(* Logix 5000 project; controller CIP_14485201 vendor 1 type 14 code 216 rev 38.11; software revision 38.01 *)

TASK MainProgram (periodic, rate 20 ms, priority 1, watchdog 40 ms) : MainProgram
TASK PID_SupplyFlow (periodic, rate 250 ms, priority 5, watchdog 500 ms) : PID_SupplyFlow

MODULES
   Local : vendor 1 type 14 code 216 (5069 0, rev 38.11)
        Module:7:I.1   // SPARE IN-426
        Module:7:I.6   // SPARE IN-436
        Module:7:I.7   // SPARE IN-438
        Module:7:I.0   // CHEM #1 TANK LOW LEVEL LSL-201
        Module:7:I.2   // CHEM #2 TANK LOW LEVEL LSL-301
        Module:7:I.3   // SPARE IN-430
        Module:7:I.4   // SPARE IN-432
        Module:7:I.5   // SPARE IN-434
        Module:7:I   // 8-PT DIG. INPUT
        Module:9:O.7   // SPARE OUT-396
        Module:9:O.0   // AIR BLOW BLOCK XY-008
        Module:9:O.2   // CHEM #1 ENABLE XY-202
        Module:9:O.3   // CHEM #2 ENABLE XY-302
        Module:9:O.5   // CHEM #2 BLOCK XY-305
        Module:9:O.6   // OVERFLOW TANK DRAIN PUMP XV-032
        Module:9:O.4   // CHEM #1 BLOCK XY-205
        Module:9:O.1   // SPARE OUT-384
        Module:9:O   // 8-PT DIG. OUTPUT
        Module:10:I   // 8-PT DIG. OUTPUT
        Module:10:O.1   // LOW POINT DRAIN XY-023
        Module:10:O.3   // SPARE SOLENOID SV-410
        Module:10:O.4   // SPARE SOLENOID SV-412
        Module:10:O.0   // OVERFLOW TANK DRAIN XY-022
        Module:10:O.2   // DRAIN TO WASTE NEUTRALIZATION XY-024
        Module:10:O.5   // SPARE OUT-414
        Module:10:O.6   // SPARE OUT-416
        Module:10:O.7   // SPARE OUT-418
        Module:10:O   // 8-PT DIG. OUTPUT
        Module:6:I.7   // SPARE IN-356
        Module:6:I.0   // SEP. TANK HIGH LEVEL LSH-101
        Module:6:I.1   // SUPPLY PUMP FAULT CONTACT JY-001C
        Module:6:I.2   // SEP. TANK MIDDLE LEVEL LSM-110
        Module:6:I.3   // HEATER CONTACTOR ALARM CONTACT JY-004B
        Module:6:I.4   // HEATER HIGH TEMP CONTACT TSH-004
        Module:6:I.5   // DRAIN PUMP LOW LEVEL LSL-405
        Module:6:I.6   // OVERFLOW TANK HIGH LEVEL LSH-401
        Module:6:I   // 8-PT DIG. INPUT
        Module:5:I.5   // SPARE IN-334
        Module:5:I.6   // SPARE IN-336
        Module:5:I.0   // CONTROL POWER ON CP-153
        Module:5:I.1   // LOCAL E-STOP PRESSED PBLT-125
        Module:5:I.2   // SEPARATOR TANK BURST SENSOR PSH-106
        Module:5:I.3   // AIR SUPPLY PRESSURE PSL-021
        Module:5:I.4   // SUPPLY PUMP AUX CONTACT JY-001B
        Module:5:I.7   // SEP. TANK LOW LEVEL LSL-105
        Module:5:I   // 8-PT DIG. INPUT
        Module:8:O.1   // AIR BLOW XV-008A
        Module:8:O.6   // ALARM HORN AH-376
        Module:8:O.5   // RETURN TO DRAIN XY-018
        Module:8:O.4   // SPARE SOLENOID SV-372
        Module:8:O.7   // HEATER ENABLE JY-004A
        Module:8:O.0   // SEP. TANK AWFI FILL XY-102
        Module:8:O.2   // SUPPLY PUMP CASING DRAIN XY-002
        Module:8:O.3   // SUPPLY PUMP ENABLE JY-001A
        Module:8:O   // 8-PT DIG. OUTPUT
        Module:8:I   // 8-PT DIG. OUTPUT
        Module:9:I.4   // SPARE IN-432
        Module:9:I.5   // SPARE IN-434
        Module:9:I.6   // SPARE IN-436
        Module:9:I.7   // SPARE IN-438
        Module:9:I.0   // CHEM 1 TANK LOW LEVEL LSL-201
        Module:9:I.1   // CHEM 1 TANK HIGH LEVEL LSH-201
        Module:9:I.2   // CHEM 2 TANK LOW LEVEL LSL-301
        Module:9:I.3   // CHEM 2 TANK HIGH LEVEL LSH-301
        Module:9:I   // 8-PT DIG. OUTPUT
      Module : 1734-AENT (Ethernet 192.168.1.50, rev 4.1, Output RPI 20 ms)
         Analog_In1 : vendor 1 type 115 code 210 (PointIO 1, rev 3.1, Input RPI 80 ms)
              Module:1:C   // 8-PT ANALOG INPUT
              Module:1:I.Ch2Data   // RINSE CONDUCTIVITY 0-10 uS/cm AE-019
              Module:1:I.Ch3Data   // WASH CONDUCTIVITY 0-100 mS/cm AE-104
              Module:1:I.Ch0Data   // SUPPLY TEMPERATURE 0-100°C TT-005
              Module:1:I.Ch1Data   // RETURN TEMPERATURE 0-100°C TT-017
              Module:1:I.Ch2Fault   // RINSE CONDUCTIVITY 0-10 uS/cm AE-019 FAULT
              Module:1:I.Ch2Underrange   // RINSE CONDUCTIVITY 0-10 uS/cm AE-019 UNDERRANGE
              Module:1:I.Ch1Underrange   // RETURN TEMPERATURE 0-100°C TT-017 UNDERRANGE
              Module:1:I.Ch1Overrange   // RETURN TEMPERATURE 0-100°C TT-017 OVERRANGE
              Module:1:I.Ch0Overrange   // SUPPLY TEMPERATURE 0-100°C TT-005 OVERRANGE
              Module:1:I.Ch1Fault   // RETURN TEMPERATURE 0-100°C TT-017 FAULT
              Module:1:I.Ch6Data   // SUPPLY PRESSURE 0-100 PSIG PIT-009
              Module:1:I.Ch7Data   // SPARE IN-272
              Module:1:I.Ch4Data   // SUPPLY FLOW 0-60 GPM FIT-010
              Module:1:I.Ch5Data   // SPARE IN-264
              Module:1:I.Ch0Fault   // SUPPLY TEMPERATURE 0-100°C TT-005 FAULT
              Module:1:I.Ch0Underrange   // SUPPLY TEMPERATURE 0-100°C TT-005 UNDERRANGE
              Module:1:I.Ch2Overrange   // RINSE CONDUCTIVITY 0-10 uS/cm AE-019 OVERRANGE
              Module:1:I.Ch3Fault   // WASH CONDUCTIVITY 0-100 mS/cm AE-104 FAULT
              Module:1:I.Ch3Underrange   // WASH CONDUCTIVITY 0-100 mS/cm AE-104 UNDERRANGE
              Module:1:I.Ch3Overrange   // WASH CONDUCTIVITY 0-100 mS/cm AE-104 OVERRANGE
              Module:1:I.Ch4Fault   // SUPPLY FLOW 0-60 GPM FIT-010 FAULT
              Module:1:I.Ch4Underrange   // SUPPLY FLOW 0-60 GPM FIT-010 UNDERRANGE
              Module:1:I.Ch4Overrange   // SUPPLY FLOW 0-60 GPM FIT-010 OVERRANGE
              Module:1:I.Ch5Fault   // SPARE IN-264 FAULT
              Module:1:I.Ch5Underrange   // SPARE IN-264 UNDERRANGE
              Module:1:I.Ch5Overrange   // SPARE IN-264 OVERRANGE
              Module:1:I.Ch6Fault   // SUPPLY PRESSURE 0-100 PSIG PIT-009 FAULT
              Module:1:I.Ch6Underrange   // SUPPLY PRESSURE 0-100 PSIG PIT-009 UNDERRANGE
              Module:1:I.Ch6Overrange   // SUPPLY PRESSURE 0-100 PSIG PIT-009 OVERRANGE
              Module:1:I.Ch7Fault   // SPARE IN-272 FAULT
              Module:1:I.Ch7Underrange   // SPARE IN-272 UNDERRANGE
              Module:1:I.Ch7Overrange   // SPARE IN-272 OVERRANGE
              Module:1:I   // 8-PT ANALOG INPUT
         Analog_In2 : 1734-IE2C (PointIO 2, rev 3.1, Input RPI 80 ms)
              Module:2:C   // 2-PT ANALOG OUTPUT
              Module:2:I.Ch1Fault   // DRAIN FLOW FEEDBACK POSTION 0-100% FY-006B FAULT
              Module:2:I.Ch1Overrange   // DRAIN FLOW FEEDBACK POSTION 0-100% FY-006B OVERRANGE
              Module:2:I.Ch0Fault   // SUPPLY FLOW FEEDBACK POSTION 0-100% FY-003B FAULT
              Module:2:I.Ch0Overrange   // SUPPLY FLOW FEEDBACK POSTION 0-100% FY-003B OVERRANGE
              Module:2:I.Ch0Underrange   // SUPPLY FLOW FEEDBACK POSTION 0-100% FY-003B UNDERRANGE
              Module:2:I.Ch1Underrange   // DRAIN FLOW FEEDBACK POSTION 0-100% FY-006B UNDERRANGE
              Module:2:I.Ch0Data   // SUPPLY FLOW FEEDBACK POSTION 0-100% FY-003B
              Module:2:I.Ch1Data   // DRAIN FLOW FEEDBACK POSTION 0-100% FY-006B
              Module:2:I   // 2-PT ANALOG OUTPUT
         Discrete_In3 : 1734-IB8 (PointIO 7, rev 3.1)
              Module:7:C   // 8-PT DIG. INPUT
         Discrete_In1 : 1734-IB8 (PointIO 5, rev 3.1)
              Module:5:C   // 8-PT DIG. INPUT
         Discrete_In2 : 1734-IB8 (PointIO 6, rev 3.1)
              Module:6:C   // 8-PT DIG. INPUT
         Discrete_Out2 : 1734-OB8 (PointIO 9, rev 3.1)
              Module:9:C   // 8-PT DIG. OUTPUT
         Analog_Out1 : 1734-OE2C (PointIO 3, rev 3.1, Output RPI 80 ms)
              Module:3:C   // 2-PT ANALOG OUTPUT
              Module:3:I.Ch0Fault   // SUPPLY FLOW FEEDBACK POSTION 0-100% FY-003B FAULT
              Module:3:I.Ch1Fault   // DRAIN FLOW FEEDBACK POSTION 0-100% FY-006B FAULT
              Module:3:I   // 2-PT ANALOG OUTPUT
              Module:3:O.Ch0Data   // SPARE OUT-284
              Module:3:O.Ch1Data   // SUPPLY FLOW MODULATION 0-100% FY-003A
              Module:3:O   // 2-PT ANALOG OUTPUT
         Analog_Out2 : 1734-OE2C (PointIO 4, rev 3.1, Output RPI 80 ms)
              Module:4:C   // 8-PT DIG. INPUT
              Module:4:I   // 8-PT DIG. INPUT
              Module:4:O.Ch0Data   // DRAIN FLOW MODULATION 0-100% FY-006A
              Module:4:O.Ch1Data   // SPARE OUT-298
              Module:4:O   // 2-PT ANALOG OUTPUT
         Discrete_Out1 : 1734-OB8 (PointIO 8, rev 3.1)
              Module:8:C   // 8-PT DIG. OUTPUT
         Discrete_Out3 : 1734-OB8 (PointIO 10, rev 3.1)
              Module:10:C   // 8-PT DIG. OUTPUT
END_MODULES

TYPE CIP_to_Process :
STRUCT
   DINT : DINT[4];
   REAL : REAL[20];
   STRING : STRING[5];
END_STRUCT
END_TYPE

TYPE Process_to_CIP :
STRUCT
   DINT : DINT[2];
   REAL : REAL[2];
END_STRUCT
END_TYPE

TYPE RECIPE :
STRUCT
   OpCode : DINT[97];   // OPCODES
   StepTime : DINT[97];   // STEP TIMES
   Setpoint : REAL[97];   // SETPOINTS
   Name : STRING;   // NAME
END_STRUCT
END_TYPE

TYPE Wash_Control :
STRUCT
   Print_Control : DINT;   // PRINT CONTROL
   Print_Control_One_Shot : DINT;   // ONE SHOT
   Print_Control_String : STRING[3];   // PRINT CONTROL STRING
   Timer : TIMER[4];   // PRINT RATE TO ASCII PORT
END_STRUCT
END_TYPE

TYPE Wash_Data :
STRUCT
   Start_Time : STRING;   // START TIME
   Stop_Time : STRING;   // STOP TIME
   Required_Time : DINT[6];   // REQUIRED TIME
   Required_Time_String : STRING[6];   // REQUIRED TIME STRING
   Temperature : DINT[3];   // TEMPERATURE
   Temperature_String : STRING[6];   // TEMPERATURE STRING
   Conductivity : DINT[3];   // CONDUCTIVITY
   Conductivity_String : STRING[6];   // CONDUCTIVITY STRING
   Flow : DINT[3];   // SUPPLY FLOW
   Flow_String : STRING[6];   // SUPPLY FLOW STRING
   Pressure : DINT[3];   // SUPPLY PRESSURE
   Pressure_String : STRING[6];   // SUPPLY PRESSURE STRING
   Sample_Timer : TIMER;   // SAMPLE TIMER
   Counter : COUNTER;   // SAMPLE COUNTER
   Print_Text : STRING[3];   // PRINT SPACE
   Active : BOOL[32];   // ACTIVE
END_STRUCT
END_TYPE

TYPE Wash_Data_Control :
STRUCT
   Control : DINT[2];   // DATA CONTROL
   One_Shot : DINT;   // DATA CONTROL ONE SHOT
   Print_Active_Pin : BOOL;   // PRINT ACTIVE PIN FROM OPCODE PINNING CHART
   Timer : TIMER;   // PRINT WASH DELAY CLEAR ALLOW FOR DATA TO BE TRANSFERED TO THE TABLE
END_STRUCT
END_TYPE

TYPE Wash_Steps :
STRUCT
   Wash_Steps : STRING[40];
   Print_Step : DINT[2];
END_STRUCT
END_TYPE

VAR_GLOBAL   (* controller tags *)
   Alarm_Ack : INT[8];   // ALARMS ACKNOWLEDGE BITS
        [2].15   // ALARM 47 ACKNOWLEDGE
        [2].2   // ALARM 34 ACKNOWLEDGE
        [2].13   // ALARM 45 ACKNOWLEDGE
        [2].14   // ALARM 46 ACKNOWLEDGE
        [6].0   // ALARM 96 ACKNOWLEDGE
        [6].1   // ALARM 97 ACKNOWLEDGE
        [6].2   // ALARM 98 ACKNOWLEDGE
        [6].10   // ALARM 106 ACKNOWLEDGE
        [6].11   // ALARM 107 ACKNOWLEDGE
        [6].12   // ALARM 108 ACKNOWLEDGE
        [6].13   // ALARM 109 ACKNOWLEDGE
        [2].3   // ALARM 35 ACKNOWLEDGE
        [2].4   // ALARM 36 ACKNOWLEDGE
        [2].5   // ALARM 37 ACKNOWLEDGE
        [6].14   // ALARM 110 ACKNOWLEDGE
        [6].15   // ALARM 111 ACKNOWLEDGE
        [2].6   // ALARM 38 ACKNOWLEDGE
        [2].7   // ALARM 39 ACKNOWLEDGE
        [2].8   // ALARM 40 ACKNOWLEDGE
        [6].3   // ALARM 99 ACKNOWLEDGE
        [6].4   // ALARM 100 ACKNOWLEDGE
        [6].5   // ALARM 101 ACKNOWLEDGE
        [2].9   // ALARM 41 ACKNOWLEDGE
        [3]   // ALARMS 48-63 ACKNOWLEDGE BITS
        [6].6   // ALARM 102 ACKNOWLEDGE
        [6].7   // ALARM 103 ACKNOWLEDGE
        [6].8   // ALARM 104 ACKNOWLEDGE
        [3].0   // ALARM 48 ACKNOWLEDGE
        [3].1   // ALARM 49 ACKNOWLEDGE
        [3].2   // ALARM 50 ACKNOWLEDGE
        [6].9   // ALARM 105 ACKNOWLEDGE
        [7]   // ALARMS 97-127 ACKNOWLEDGE BITS
        [3].10   // ALARM 58 ACKNOWLEDGE
        [3].11   // ALARM 59 ACKNOWLEDGE
        [0]   // ALARMS 1-15 ACKNOWLEDGE BITS
        [7].0   // ALARM 112 ACKNOWLEDGE
        [7].1   // ALARM 113 ACKNOWLEDGE
        [7].10   // ALARM 122 ACKNOWLEDGE
        [3].12   // ALARM 60 ACKNOWLEDGE
        [3].13   // ALARM 61 ACKNOWLEDGE
        [0].1   // ALARM 1 ACKNOWLEDGE
        [0].10   // ALARM 10 ACKNOWLEDGE
        [7].11   // ALARM 123 ACKNOWLEDGE
        [7].12   // ALARM 124 ACKNOWLEDGE
        [3].14   // ALARM 62 ACKNOWLEDGE
        [3].15   // ALARM 63 ACKNOWLEDGE
        [0].11   // ALARM 11 ACKNOWLEDGE
        [0].12   // ALARM 12 ACKNOWLEDGE
        [7].13   // ALARM 125 ACKNOWLEDGE
        [7].14   // ALARM 126 ACKNOWLEDGE
        [3].3   // ALARM 51 ACKNOWLEDGE
        [3].4   // ALARM 52 ACKNOWLEDGE
        [3].5   // ALARM 53 ACKNOWLEDGE
        [0].13   // ALARM 13 ACKNOWLEDGE
        [0].14   // ALARM 14 ACKNOWLEDGE
        [7].15   // ALARM 127 ACKNOWLEDGE
        [7].2   // ALARM 114 ACKNOWLEDGE
        [7].3   // ALARM 115 ACKNOWLEDGE
        [3].6   // ALARM 54 ACKNOWLEDGE
        [3].7   // ALARM 55 ACKNOWLEDGE
        [3].8   // ALARM 56 ACKNOWLEDGE
        [0].15   // ALARM 15 ACKNOWLEDGE
        [0].2   // ALARM 2 ACKNOWLEDGE
        [7].4   // ALARM 116 ACKNOWLEDGE
        [7].5   // ALARM 117 ACKNOWLEDGE
        [7].6   // ALARM 118 ACKNOWLEDGE
        [3].9   // ALARM 57 ACKNOWLEDGE
        [4]   // ALARMS 64-79 ACKNOWLEDGE BITS
        [0].3   // ALARM 3 ACKNOWLEDGE
        [0].4   // ALARM 4 ACKNOWLEDGE
        [0].5   // ALARM 5 ACKNOWLEDGE
        [7].7   // ALARM 119 ACKNOWLEDGE
        [7].8   // ALARM 120 ACKNOWLEDGE
        [7].9   // ALARM 121 ACKNOWLEDGE
        [4].0   // ALARM 64 ACKNOWLEDGE
        [4].1   // ALARM 65 ACKNOWLEDGE
        [4].2   // ALARM 66 ACKNOWLEDGE
        [0].6   // ALARM 6 ACKNOWLEDGE
        [0].7   // ALARM 7 ACKNOWLEDGE
        [0].8   // ALARM 8 ACKNOWLEDGE
        [4].10   // ALARM 74 ACKNOWLEDGE
        [4].11   // ALARM 75 ACKNOWLEDGE
        [0].9   // ALARM 9 ACKNOWLEDGE
        [1]   // ALARMS 16-31 ACKNOWLEDGE BITS
        [4].12   // ALARM 76 ACKNOWLEDGE
        [4].13   // ALARM 77 ACKNOWLEDGE
        [1].0   // ALARM 16 ACKNOWLEDGE
        [1].1   // ALARM 17 ACKNOWLEDGE
        [4].14   // ALARM 78 ACKNOWLEDGE
        [4].15   // ALARM 79 ACKNOWLEDGE
        [1].10   // ALARM 26 ACKNOWLEDGE
        [1].11   // ALARM 27 ACKNOWLEDGE
        [4].3   // ALARM 67 ACKNOWLEDGE
        [4].4   // ALARM 68 ACKNOWLEDGE
        [4].5   // ALARM 69 ACKNOWLEDGE
        [1].12   // ALARM 28 ACKNOWLEDGE
        [1].13   // ALARM 29 ACKNOWLEDGE
        [4].6   // ALARM 70 ACKNOWLEDGE
        [4].7   // ALARM 71 ACKNOWLEDGE
        [4].8   // ALARM 72 ACKNOWLEDGE
        [1].14   // ALARM 30 ACKNOWLEDGE
        [1].15   // ALARM 31 ACKNOWLEDGE
        [4].9   // ALARM 73 ACKNOWLEDGE
        [5]   // ALARMS 80-95 ACKNOWLEDGE BITS
        [1].2   // ALARM 18 ACKNOWLEDGE
        [1].3   // ALARM 19 ACKNOWLEDGE
        [5].0   // ALARM 80 ACKNOWLEDGE
        [5].1   // ALARM 81 ACKNOWLEDGE
        [5].2   // ALARM 82 ACKNOWLEDGE
        [1].4   // ALARM 20 ACKNOWLEDGE
        [1].5   // ALARM 21 ACKNOWLEDGE
        [5].10   // ALARM 90 ACKNOWLEDGE
        [5].11   // ALARM 91 ACKNOWLEDGE
        [1].6   // ALARM 22 ACKNOWLEDGE
        [1].7   // ALARM 23 ACKNOWLEDGE
        [5].12   // ALARM 92 ACKNOWLEDGE
        [5].13   // ALARM 93 ACKNOWLEDGE
        [1].8   // ALARM 24 ACKNOWLEDGE
        [1].9   // ALARM 25 ACKNOWLEDGE
        [5].14   // ALARM 94 ACKNOWLEDGE
        [5].15   // ALARM 95 ACKNOWLEDGE
        [2]   // ALARMS 32-47 ACKNOWLEDGE BITS
        [2].0   // ALARM 32 ACKNOWLEDGE
        [5].3   // ALARM 83 ACKNOWLEDGE
        [5].4   // ALARM 84 ACKNOWLEDGE
        [5].5   // ALARM 85 ACKNOWLEDGE
        [2].1   // ALARM 33 ACKNOWLEDGE
        [2].10   // ALARM 42 ACKNOWLEDGE
        [5].6   // ALARM 86 ACKNOWLEDGE
        [5].7   // ALARM 87 ACKNOWLEDGE
        [5].8   // ALARM 88 ACKNOWLEDGE
        [2].11   // ALARM 43 ACKNOWLEDGE
        [2].12   // ALARM 44 ACKNOWLEDGE
        [5].9   // ALARM 89 ACKNOWLEDGE
        [6]   // ALARMS 96-111 ACKNOWLEDGE BITS
   Alarm_Ack_All_PB : BOOL;   // SYSTEM ALARM ACK ALL PUSHBUTTON ON ALARM PAGE
   Alarm_Present : INT[8] := ([0] := 70, [2] := 98);   // ALARM MSGS 1-127 PRESENT BITS
        [7].0   // ALARM 112 PRESENT
        [7].1   // ALARM 113 PRESENT
        [7].10   // ALARM 122 PRESENT
        [1].3   // ALARM 19 SUPPLY TEMPERATURE HOLD WATCHDOG PRESENT
        [1].4   // ALARM 20 RETURN TEMPERATURE HOLD WATCHDOG PRESENT
        [1].15   // ALARM 31 SEPARATOR TANK LOW LEVEL PRESENT
        [1].2   // ALARM 18 SEPARATOR TANK EMPTY HOLD WATCHDOG PRESENT
        [7].11   // ALARM 123 PRESENT
        [7].12   // ALARM 124 PRESENT
        [7].13   // ALARM 125 PRESENT
        [3].0   // ALARM 48 PRESENT
        [3].1   // ALARM 49 PRESENT
        [3].10   // ALARM 58 PRESENT
        [7].14   // ALARM 126 PRESENT
        [7].15   // ALARM 127 PRESENT
        [7].2   // ALARM 114 PRESENT
        [3].11   // ALARM 59 PRESENT
        [3].12   // ALARM 60 PRESENT
        [3].13   // ALARM 61 PRESENT
        [7].3   // ALARM 115 PRESENT
        [7].4   // ALARM 116 PRESENT
        [7].5   // ALARM 117 PRESENT
        [3].14   // ALARM 62 PRESENT
        [3].15   // ALARM 63 PRESENT
        [3].2   // ALARM 50 PRESENT
        [7].6   // ALARM 118 PRESENT
        [7].7   // ALARM 119 PRESENT
        [7].8   // ALARM 120 PRESENT
        [3].3   // ALARM 51 PRESENT
        [3].4   // ALARM 52 PRESENT
        [3].5   // ALARM 53 PRESENT
        [7].9   // ALARM 121 PRESENT
        [3].6   // ALARM 54 PRESENT
        [3].7   // ALARM 55 PRESENT
        [3].8   // ALARM 56 PRESENT
        [3].9   // ALARM 57 PRESENT
        [4]   // ALARM MSGS 64-79 PRESENT BITS
        [4].0   // ALARM 64 PRESENT
        [4].1   // ALARM 65 PRESENT
        [4].10   // ALARM 74 PRESENT
        [4].11   // ALARM 75 PRESENT
        [4].12   // ALARM 76 PRESENT
        [4].13   // ALARM 77 PRESENT
        [4].14   // ALARM 78 PRESENT
        [4].15   // ALARM 79 PRESENT
        [4].2   // ALARM 66 PRESENT
        [4].3   // ALARM 67 PRESENT
        [4].4   // ALARM 68 PRESENT
        [4].5   // ALARM 69 PRESENT
        [4].6   // ALARM 70 PRESENT
        [4].7   // ALARM 71 PRESENT
        [4].8   // ALARM 72 PRESENT
        [4].9   // ALARM 73 PRESENT
        [5]   // ALARM MSGS 80-95 PRESENT BITS
        [5].0   // ALARM 80 PRESENT
        [5].1   // ALARM 81 PRESENT
        [5].10   // ALARM 90 PRESENT
        [5].11   // ALARM 91 PRESENT
        [5].12   // ALARM 92 PRESENT
        [5].13   // ALARM 93 PRESENT
        [0]   // ALARM MSGS 1-15 PRESENT BITS
        [0].0   // ALARM 0 N/A PRESENT
        [5].14   // ALARM 94 PRESENT
        [5].15   // ALARM 95 PRESENT
        [5].2   // ALARM 82 PRESENT
        [0].1   // ALARM 1 LOSS OF CONTROL POWER PRESENT
        [0].10   // ALARM 10 WASH CONDUCTIVITY SENSOR FAILURE PRESENT
        [0].5   // ALARM 5 PRESENT
        [5].3   // ALARM 83 PRESENT
        [5].4   // ALARM 84 PRESENT
        [5].5   // ALARM 85 PRESENT
        [0].11   // ALARM 11 SUPPLY FLOW SENSOR FAILURE PRESENT
        [0].12   // ALARM 12 SUPPLY FLOW FEEDBACK SENSOR FAILURE PRESENT
        [5].6   // ALARM 86 PRESENT
        [5].7   // ALARM 87 PRESENT
        [5].8   // ALARM 88 PRESENT
        [0].13   // ALARM 13 SUPPLY PRESSURE SENSOR FAILURE PRESENT
        [0].14   // ALARM 14 DRAIN FLOW FEEDBACK SENSOR FAILURE PRESENT
        [5].9   // ALARM 89 PRESENT
        [6]   // ALARM MSGS 96-111 PRESENT BITS
        [0].15   // ALARM 15 SUPPLY PUMP FAILURE PRESENT
        [0].2   // ALARM 2 LOSS OF PLC POWER PRESENT
        [6].0   // ALARM 96 PRESENT
        [6].1   // ALARM 97 PRESENT
        [6].10   // ALARM 106 PRESENT
        [0].3   // ALARM 3 LOCAL E-STOP PRESSED PRESENT
        [0].6   // ALARM 6 I/O COMMUNICATION FAILURE PRESENT
        [0].4   // ALARM 4 PRESENT
        [1].5   // ALARM 21 RINSE CONDUCTIVITY HOLD WATCHDOG PRESENT
        [1].6   // ALARM 22 CHEM #1 CONDUCTIVITY HOLD WATCHDOG PRESENT
        [6].11   // ALARM 107 PRESENT
        [6].12   // ALARM 108 PRESENT
        [6].2   // ALARM 98 PRESENT
        [0].7   // ALARM 7 SUPPLY TEMPERATURE SENSOR FAILURE PRESENT
        [0].8   // ALARM 8 RETURN TEMPERATURE SENSOR FAILURE PRESENT
        [1].7   // ALARM 23 CHEM #2 CONDUCTIVITY HOLD WATCHDOG PRESENT
        [1].8   // ALARM 24 OVERFLOW TANK EMPTY HOLD WATCHDOG PRESENT
        [6].13   // ALARM 109 PRESENT
        [6].14   // ALARM 110 PRESENT
        [6].3   // ALARM 99 PRESENT
        [0].9   // ALARM 9 RINSE CONDUCTIVITY SENSOR FAILURE PRESENT
        [1]   // ALARM MSGS 16-31 PRESENT BITS
        [6].15   // ALARM 111 PRESENT
        [6].4   // ALARM 100 PRESENT
        [6].5   // ALARM 101 PRESENT
        [1].1   // ALARM 17 SEPARATOR TANK FILL HOLD WATCHDOG PRESENT
        [1].10   // ALARM 26 HIGH SUPPLY FLOW PRESENT
        [6].6   // ALARM 102 PRESENT
        [6].7   // ALARM 103 PRESENT
        [6].8   // ALARM 104 PRESENT
        [1].11   // ALARM 27 LOW SUPPLY FLOW PRESENT
        [1].12   // ALARM 28 HIGH SUPPLY PRESSURE PRESENT
        [1].0   // ALARM 16 PRESENT
        [6].9   // ALARM 105 PRESENT
        [7]   // ALARM MSGS 112-127 PRESENT BITS
        [1].13   // ALARM 29 LOW SUPPLY PRESSURE PRESENT
        [1].14   // ALARM 30 PRESENT
        [2].0   // ALARM 32 PRESENT
        [1].9   // ALARM 25 HIGH SUPPLY TEMPERATURE PRESENT
        [2]   // ALARM MSGS 32-47 PRESENT BITS
        [2].1   // ALARM 33 HEATER CONTACTOR FAULT PRESENT
        [2].10   // ALARM 42 PRESENT
        [2].11   // ALARM 43 PRESENT
        [2].12   // ALARM 44 PRESENT
        [2].13   // ALARM 45 PRESENT
        [2].14   // ALARM 46 PROCESS EQUIPMENT HEARTBEAT FAILURE PRESENT
        [2].15   // ALARM 47 PROCESS EQUIPMENT STOP ACTIVE PRESENT
        [2].2   // ALARM 34 HEATER ELEMENT HIGH TEMPERATURE PRESENT
        [2].3   // ALARM 35 CHEM #1 TANK LOW LEVEL PRESENT
        [2].4   // ALARM 36 CHEM #2 TANK LOW LEVEL PRESENT
        [2].5   // ALARM 37 PANEL AIR PRESSURE FAILURE PRESENT
        [2].6   // ALARM 38 SEP. TANK BURST SENSOR FAILURE PRESENT
        [2].8   // ALARM 40 SUPPLY FLOW MODULATION VALVE FAILURE PRESENT
        [2].9   // ALARM 41 DRAIN FLOW MODULATION VALVE FAILURE PRESENT
        [3]   // ALARM MSGS 48-63 PRESENT BITS
        [2].7   // ALARM 39 PRESENT
   Alarm_Preset_Indx : DINT := 84;   // ALARM TIMER PRESET INDEX POSITION
   Alarm_Remote_Ack_All : BOOL;   // SYSTEM ALARM ACK ALL TAG USED ON ALARM SETUP ADVANCED TAB TOGGLES EVEYTIME THE ACK_ALL BUTTON IS PUSHED
   Alarm_Status_Reset : BOOL;   // SYSTEM ALARM ACK ALL TAG USED ON ALARM SETUP ADVANCED TAB TOGGLES EVERYTIME THE HISTORY CLEAR ALL IS PUSHED
   Alarm_Timer : TIMER[128] := ([1].ACC := 20, [1].EN := 1, [1].DN := 1, [2].ACC := 20, [2].EN := 1, [2].DN := 1, [6].PRE := 3000, [7].PRE := 5000, [8].PRE := 5000, [9].PRE := 5000, [10].PRE := 5000, [11].PRE := 5000, [12].PRE := 5000, [13].PRE := 5000, [14].PRE := 5000, [15].PRE := 3000, [17].PRE := 180000, [18].PRE := 180000, [19].PRE := 300000, [20].PRE := 900000, [21].PRE := 900000, [22].PRE := 300000, [23].PRE := 300000, [24].PRE := 300000, [25].PRE := 1000, [26].PRE := 8000, [27].PRE := 15000, [28].PRE := 5000, [29].PRE := 15000, [33].PRE := 3000, [34].PRE := 3000, [35].PRE := 500, [36].PRE := 500, [37].PRE := 3000, [38].ACC := 20, [38].EN := 1, [38].DN := 1, [39].ACC := 20, [39].EN := 1, [39].DN := 1, [40].PRE := 10000, [41].PRE := 10000, [42].ACC := 20, [42].EN := 1, [42].DN := 1, [43].PRE := 1000, [43].ACC := 1000, [43].EN := 1, [43].DN := 1, [44].PRE := 1000, [45].ACC := 20, [45].EN := 1, [45].DN := 1, [46].PRE := 10000, [48].ACC := 20, [48].EN := 1, [48].DN := 1, [49].ACC := 20, [49].EN := 1, [49].DN := 1,
        [50].ACC := 20, [50].EN := 1, [50].DN := 1, [51].ACC := 20, [51].EN := 1, [51].DN := 1, [52].ACC := 20, [52].EN := 1, [52].DN := 1, [53].ACC := 20, [53].EN := 1, [53].DN := 1, [54].ACC := 20, [54].EN := 1, [54].DN := 1, [55].ACC := 20, [55].EN := 1, [55].DN := 1, [56].ACC := 20, [56].EN := 1, [56].DN := 1, [57].ACC := 20, [57].EN := 1, [57].DN := 1, [58].ACC := 20, [58].EN := 1, [58].DN := 1, [59].ACC := 20, [59].EN := 1, [59].DN := 1, [60].ACC := 20, [60].EN := 1, [60].DN := 1, [61].ACC := 20, [61].EN := 1, [61].DN := 1, [62].ACC := 20, [62].EN := 1, [62].DN := 1, [63].ACC := 20, [63].EN := 1, [63].DN := 1, [64].ACC := 20, [64].EN := 1, [64].DN := 1, [65].ACC := 20, [65].EN := 1, [65].DN := 1, [66].ACC := 20, [66].EN := 1, [66].DN := 1, [67].ACC := 20, [67].EN := 1, [67].DN := 1, [68].ACC := 20, [68].EN := 1, [68].DN := 1, [69].ACC := 20, [69].EN := 1, [69].DN := 1,
        [70].ACC := 20, [70].EN := 1, [70].DN := 1, [71].ACC := 20, [71].EN := 1, [71].DN := 1, [72].ACC := 20, [72].EN := 1, [72].DN := 1, [73].ACC := 20, [73].EN := 1, [73].DN := 1, [74].ACC := 20, [74].EN := 1, [74].DN := 1, [75].ACC := 20, [75].EN := 1, [75].DN := 1, [76].ACC := 20, [76].EN := 1, [76].DN := 1, [77].ACC := 20, [77].EN := 1, [77].DN := 1, [78].ACC := 20, [78].EN := 1, [78].DN := 1, [79].ACC := 20, [79].EN := 1, [79].DN := 1, [80].ACC := 20, [80].EN := 1, [80].DN := 1, [81].ACC := 20, [81].EN := 1, [81].DN := 1, [82].ACC := 20, [82].EN := 1, [82].DN := 1, [83].ACC := 20, [83].EN := 1, [83].DN := 1, [84].ACC := 20, [84].EN := 1, [84].DN := 1, [85].ACC := 20, [85].EN := 1, [85].DN := 1, [86].ACC := 20, [86].EN := 1, [86].DN := 1, [87].ACC := 20, [87].EN := 1, [87].DN := 1, [88].ACC := 20, [88].EN := 1, [88].DN := 1, [89].ACC := 20, [89].EN := 1, [89].DN := 1,
        [90].ACC := 20, [90].EN := 1, [90].DN := 1, [91].ACC := 20, [91].EN := 1, [91].DN := 1, [92].ACC := 20, [92].EN := 1, [92].DN := 1, [93].ACC := 20, [93].EN := 1, [93].DN := 1, [94].ACC := 20, [94].EN := 1, [94].DN := 1, [95].ACC := 20, [95].EN := 1, [95].DN := 1, [96].ACC := 20, [96].EN := 1, [96].DN := 1, [97].ACC := 20, [97].EN := 1, [97].DN := 1, [98].ACC := 20, [98].EN := 1, [98].DN := 1, [99].ACC := 20, [99].EN := 1, [99].DN := 1, [100].ACC := 20, [100].EN := 1, [100].DN := 1, [101].ACC := 20, [101].EN := 1, [101].DN := 1, [102].ACC := 20, [102].EN := 1, [102].DN := 1, [103].ACC := 20, [103].EN := 1, [103].DN := 1, [104].ACC := 20, [104].EN := 1, [104].DN := 1, [105].ACC := 20, [105].EN := 1, [105].DN := 1, [106].ACC := 20, [106].EN := 1, [106].DN := 1, [107].ACC := 20, [107].EN := 1, [107].DN := 1, [108].ACC := 20, [108].EN := 1, [108].DN := 1, [109].ACC := 20, [109].EN := 1, [109].DN := 1,
        [110].ACC := 20, [110].EN := 1, [110].DN := 1, [111].ACC := 20, [111].EN := 1, [111].DN := 1, [112].ACC := 20, [112].EN := 1, [112].DN := 1, [113].ACC := 20, [113].EN := 1, [113].DN := 1, [114].ACC := 20, [114].EN := 1, [114].DN := 1, [115].ACC := 20, [115].EN := 1, [115].DN := 1, [116].ACC := 20, [116].EN := 1, [116].DN := 1, [117].ACC := 20, [117].EN := 1, [117].DN := 1, [118].ACC := 20, [118].EN := 1, [118].DN := 1, [119].ACC := 20, [119].EN := 1, [119].DN := 1, [120].ACC := 20, [120].EN := 1, [120].DN := 1, [121].ACC := 20, [121].EN := 1, [121].DN := 1, [122].ACC := 20, [122].EN := 1, [122].DN := 1, [123].ACC := 20, [123].EN := 1, [123].DN := 1, [124].ACC := 20, [124].EN := 1, [124].DN := 1, [125].ACC := 20, [125].EN := 1, [125].DN := 1, [126].ACC := 20, [126].EN := 1, [126].DN := 1, [127].ACC := 20, [127].EN := 1, [127].DN := 1);   // ALARM MSGS 1-127 DELAY TIMERS
        [41]   // ALARM 41 DRAIN FLOW MODULATION VALVE FAILURE DELAY TIMER
        [43]   // ALARM 43 DELAY TIMER
        [44]   // ALARM 44 DELAY TIMER
        [45]   // ALARM 45 DELAY TIMER
        [0]   // ALARM 0 N/A DELAY TIMER
        [100]   // ALARM 100 DELAY TIMER
        [66]   // ALARM 66 DELAY TIMER
        [67]   // ALARM 67 DELAY TIMER
        [37]   // ALARM 37 PANEL AIR PRESSURE FAILURE DELAY TIMER
        [38]   // ALARM 38 SEP. TANK BURST SENSOR FAILURE DELAY TIMER
        [73]   // ALARM 73 DELAY TIMER
        [74]   // ALARM 74 DELAY TIMER
        [77]   // ALARM 77 DELAY TIMER
        [78]   // ALARM 78 DELAY TIMER
        [68]   // ALARM 68 DELAY TIMER
        [69]   // ALARM 69 DELAY TIMER
        [6]   // ALARM 6 I/O COMMUNICATION FAILURE DELAY TIMER
        [70]   // ALARM 70 DELAY TIMER
        [101]   // ALARM 101 DELAY TIMER
        [102]   // ALARM 102 DELAY TIMER
        [105]   // ALARM 105 DELAY TIMER
        [106]   // ALARM 106 DELAY TIMER
        [75]   // ALARM 75 DELAY TIMER
        [76]   // ALARM 76 DELAY TIMER
        [39]   // ALARM 39 DELAY TIMER
        [3]   // ALARM 3 LOCAL E-STOP PRESSED DELAY TIMER
        [80]   // ALARM 80 DELAY TIMER
        [81]   // ALARM 81 DELAY TIMER
        [71]   // ALARM 71 DELAY TIMER
        [72]   // ALARM 72 DELAY TIMER
        [103]   // ALARM 103 DELAY TIMER
        [104]   // ALARM 104 DELAY TIMER
        [40]   // ALARM 40 SUPPLY FLOW MODULATION VALVE FAILURE DELAY TIMER
        [42]   // ALARM 42 DELAY TIMER
        [79]   // ALARM 79 DELAY TIMER
        [7]   // ALARM 7 SUPPLY TEMPERATURE SENSOR FAILURE DELAY TIMER
        [82]   // ALARM 82 DELAY TIMER
        [83]   // ALARM 83 DELAY TIMER
        [107]   // ALARM 107 DELAY TIMER
        [108]   // ALARM 108 DELAY TIMER
        [84]   // ALARM 84 DELAY TIMER
        [85]   // ALARM 85 DELAY TIMER
        [109]   // ALARM 109 DELAY TIMER
        [10]   // ALARM 10 WASH CONDUCTIVITY SENSOR FAILURE DELAY TIMER
        [86]   // ALARM 86 DELAY TIMER
        [87]   // ALARM 87 DELAY TIMER
        [110]   // ALARM 110 DELAY TIMER
        [111]   // ALARM 111 DELAY TIMER
        [88]   // ALARM 88 DELAY TIMER
        [89]   // ALARM 89 DELAY TIMER
        [112]   // ALARM 112 DELAY TIMER
        [113]   // ALARM 113 DELAY TIMER
        [8]   // ALARM 8 RETURN TEMPERATURE SENSOR FAILURE DELAY TIMER
        [90]   // ALARM 90 DELAY TIMER
        [114]   // ALARM 114 DELAY TIMER
        [115]   // ALARM 115 DELAY TIMER
        [4]   // ALARM 4 DELAY TIMER
        [91]   // ALARM 91 DELAY TIMER
        [92]   // ALARM 92 DELAY TIMER
        [116]   // ALARM 116 DELAY TIMER
        [117]   // ALARM 117 DELAY TIMER
        [93]   // ALARM 93 DELAY TIMER
        [94]   // ALARM 94 DELAY TIMER
        [118]   // ALARM 118 DELAY TIMER
        [119]   // ALARM 119 DELAY TIMER
        [95]   // ALARM 95 DELAY TIMER
        [96]   // ALARM 96 DELAY TIMER
        [11]   // ALARM 11 SUPPLY FLOW SENSOR FAILURE DELAY TIMER
        [120]   // ALARM 120 DELAY TIMER
        [97]   // ALARM 97 DELAY TIMER
        [98]   // ALARM 98 DELAY TIMER
        [121]   // ALARM 121 DELAY TIMER
        [122]   // ALARM 122 DELAY TIMER
        [99]   // ALARM 99 DELAY TIMER
        [9]   // ALARM 9 RINSE CONDUCTIVITY SENSOR FAILURE DELAY TIMER
        [123]   // ALARM 123 DELAY TIMER
        [124]   // ALARM 124 DELAY TIMER
        [125]   // ALARM 125 DELAY TIMER
        [126]   // ALARM 126 DELAY TIMER
        [127]   // ALARM 127 DELAY TIMER
        [12]   // ALARM 12 SUPPLY FLOW FEEDBACK SENSOR FAILURE DELAY TIMER
        [5]   // ALARM 5 DELAY TIMER
        [13]   // ALARM 13 SUPPLY PRESSURE SENSOR FAILURE DELAY TIMER
        [16]   // ALARM 16 DELAY TIMER
        [14]   // ALARM 14 DRAIN FLOW FEEDBACK SENSOR FAILURE DELAY TIMER
        [15]   // ALARM 15 SUPPLY PUMP FAILURE DELAY TIMER
        [17]   // ALARM 17 SEPARATOR TANK FILL HOLD WATCHDOG DELAY TIMER
        [27]   // ALARM 27 LOW SUPPLY FLOW DELAY TIMER
        [18]   // ALARM 18 SEPARATOR TANK EMPTY HOLD WATCHDOG DELAY TIMER
        [1]   // ALARM 1 LOSS OF CONTROL POWER DELAY TIMER
        [19]   // ALARM 19 SUPPLY TEMPERATURE HOLD WATCHDOG DELAY TIMER
        [29]   // ALARM 29 LOW SUPPLY PRESSURE DELAY TIMER
        [20]   // ALARM 20 RETURN TEMPERATURE HOLD WATCHDOG DELAY TIMER
        [2]   // ALARM 2 LOSS OF PLC POWER DELAY TIMER
        [21]   // ALARM 21 RINSE CONDUCTIVITY HOLD WATCHDOG DELAY TIMER
        [30]   // ALARM 30 DELAY TIMER
        [46]   // ALARM 46 PROCESS EQUIPMENT HEARTBEAT FAILURE DELAY TIMER
        [48]   // ALARM 48 DELAY TIMER
        [22]   // ALARM 22 CHEM #1 CONDUCTIVITY HOLD WATCHDOG DELAY TIMER
        [25]   // ALARM 25 HIGH SUPPLY TEMPERATURE DELAY TIMER
        [47]   // ALARM 47 PROCESS EQUIPMENT STOP ACTIVE DELAY TIMER
        [49]   // ALARM 49 DELAY TIMER
        [23]   // ALARM 23 CHEM #2 CONDUCTIVITY HOLD WATCHDOG DELAY TIMER
        [26]   // ALARM 26 HIGH SUPPLY FLOW DELAY TIMER
        [24]   // ALARM 24 OVERFLOW TANK EMPTY HOLD WATCHDOG DELAY TIMER
        [28]   // ALARM 28 HIGH SUPPLY PRESSURE DELAY TIMER
        [31]   // ALARM 31 SEPARATOR TANK LOW LEVEL DELAY TIMER
        [32]   // ALARM 32 DELAY TIMER
        [33]   // ALARM 33 HEATER CONTACTOR FAULT DELAY TIMER
        [34]   // ALARM 34 HEATER ELEMENT HIGH TEMPERATURE DELAY TIMER
        [50]   // ALARM 50 DELAY TIMER
        [51]   // ALARM 51 DELAY TIMER
        [52]   // ALARM 52 DELAY TIMER
        [53]   // ALARM 53 DELAY TIMER
        [54]   // ALARM 54 DELAY TIMER
        [55]   // ALARM 55 DELAY TIMER
        [56]   // ALARM 56 DELAY TIMER
        [57]   // ALARM 57 DELAY TIMER
        [58]   // ALARM 58 DELAY TIMER
        [59]   // ALARM 59 DELAY TIMER
        [60]   // ALARM 60 DELAY TIMER
        [61]   // ALARM 61 DELAY TIMER
        [62]   // ALARM 62 DELAY TIMER
        [63]   // ALARM 63 DELAY TIMER
        [64]   // ALARM 64 DELAY TIMER
        [65]   // ALARM 65 DELAY TIMER
        [35]   // ALARM 35 CHEM #1 TANK LOW LEVEL DELAY TIMER
        [36]   // ALARM 36 CHEM #2 TANK LOW LEVEL DELAY TIMER
   Alarm_Timer_Preset : DINT[128] := ([6] := 3000, [7] := 5000, [8] := 5000, [9] := 5000, [10] := 5000, [11] := 5000, [12] := 5000, [13] := 5000, [14] := 5000, [15] := 3000, [17] := 180000, [18] := 180000, [19] := 300000, [20] := 900000, [21] := 900000, [22] := 300000, [23] := 300000, [24] := 300000, [25] := 1000, [26] := 8000, [27] := 15000, [28] := 5000, [29] := 15000, [33] := 3000, [34] := 3000, [35] := 500, [36] := 500, [37] := 3000, [40] := 10000, [41] := 10000, [43] := 1000, [44] := 1000, [46] := 10000);   // ALARM TIMER PRESETS STORAGE
   Bit : BOOL[128] := ([5] := 1, [6] := 1, [15] := 1, [16] := 1, [25] := 1, [26] := 1, [39] := 1, [40] := 1, [49] := 1, [53] := 1, [54] := 1, [62] := 1, [64] := 1, [66] := 1, [68] := 1, [77] := 1, [82] := 1, [100] := 1);   // BIT
        [0]   // SYSTEM START
        [100]   // SUPPLY TEMPERATURE CONTROL INTERLOCK
        [15]   // SUPPLY TEMPERATURE AT SETPOINT
        [20]   // CIP RUN
        [3]   // SYSTEM ABORT
        [16]   // RETURN TEMPERATURE AT SETPOINT
        [18]   // SEPARATOR LOW LEVEL RECOVERY
        [26]   // SEPARATOR TANK FILL COMPLETE
        [27]   // CHEM #1 CONDUCTIVITY AT SETPOINT
        [14]   // SYSTEM LOW LEVEL
        [21]   // CIP LATCH
        [22]   // CIP ABORT
        [9]   // DRAINS OPEN
        [48]   // SYSTEM IN LOW LEVEL RECOVERY
        [81]   // REPORT TICKET PRINTING ACTIVE START PROHIBITED
        [36]   // ONE SHOT
        [34]   // SEPARATOR FILL REQUIRED
        [40]   // SHUTDOWN ALARM EXISTS
        [43]   // CHEM #1 CONDUCTIVITY IS GREATER THAN OR EQUAL TO THE LOW HOLD LIMIT
        [7]   // OVERFLOW TANK HIGH LEVEL
        [44]   // CHEM #2 CONDUCTIVITY IS GREATER THAN OR EQUAL TO THE LOW HOLD LIMIT
        [80]   // POWER ON DWELL DONE
        [1]   // SYSTEM STOP
        [8]   // DRAIN PUMP ENABLED
        [39]   // ALARM HORN ACTIVE
        [2]   // SYSTEM HOLD
        [12]   // SYSTEM MANUAL STEP
        [17]   // RECIPE HOLD ACTIVE
        [28]   // CHEM #2 CONDUCTIVITY AT SETPOINT
        [29]   // RINSE CONDUCTIVITY AT SETPOINT
   CIP_to_Process : CIP_to_Process := (DINT[0] := 4, DINT[2] := 32, REAL[0] := 24.988554, REAL[1] := 24.843582, REAL[2] := 9.99237, REAL[6] := -1.1597742, REAL[7] := -1.1063635, STRING[2] := '0:00', STRING[3] := 'FAT TEST RECIPE');   // CIP TO PROCESS SIGNALS
        .DINT[1].1   // PBLT-125 Local E-Stop Pressed
        .REAL[1]   // TT-017 Return Temperature 0-100 deg C
        .REAL[8]   // FY-003 Supply Flow Modulation Flow Valve Output 0-100%
        .REAL[7]   // FY-006 Drain Flow Modulation Flow Valve Feedback 0-100%
        .DINT[1].2   // PSH-106 Separator Tank Burst Sensor
        .DINT[0]   // CIP DISCRETE SIGNALS
        .REAL[9]   // FY-006 Drain Flow Modulation Flow Valve Output 0-100%
        .DINT[1].8   // LSM-110 Separator Tank Middle Level
        .DINT[1].9   // JY-004B Heater Contactor Alarm Contact
        .REAL[6]   // FY-003 Supply Flow Modulation Flow Valve Feedback 0-100%
        .DINT[2].15   // XY-024 Drain to Waste Neutralization
        .DINT[0].0   // XA-099 Heartbeat to DCS
        .DINT[2].6   // JY-004A Heater Enable
        .DINT[1].11   // LSL-405 Drain Pump Low Level
        .REAL[2]   // AE-019 Rinse Conductivity 0-10 uS/cm
        .DINT[0].1   // 3CIP-3200 Skid Running
        .DINT[1].10   // TSH-004 Heater High Temp Contact
        .DINT[1].13   // LSL-201 Chem #1 Tank Low Level
        .DINT[0].2   // 3CIP-3200 Common Trouble Alarm
        .DINT[1].12   // LSH-401 Overflow Tank High Level
        .DINT[1].5   // LSL-105 Separator Tank Low Level
        .DINT[1].6   // LSH-101 Separator Tank High Level
        .DINT[1].7   // JY-001C Supply Pump Fault Contact
        .DINT[2].0   // XY-102 Separator Tank AWFI Fill
        .DINT[2].1   // XV-008A Air Blow
        .DINT[2].10   // XY-205 Chem #1 Block
        .DINT[2].11   // XY-305 Chem #2 Block
        .DINT[2].12   // XV-032 Overflow Tank Drain Pump
        .DINT[2].13   // XV-022 Overflow Tank Drain
        .DINT[2].14   // XY-023 Low Point Drain
        .DINT[2].2   // XY-002 Supply Pump Casing Drain
        .DINT[2].7   // XY-008 Air Blow Block
        .REAL[3]   // AE-104 Wash Conductivity 0-100 mS/cm
        .REAL[4]   // FIT-010 Supply Flow 0-60 gpm
        .DINT[1].14   // LSL-301 Chem #2 Tank Low Level
        .DINT[1].3   // PSL-021 Air Supply Pressure
        .DINT[2].8   // XY-202 Chem #1 Enable
        .REAL[5]   // PIT-009 Supply Pressure 0-100 psig
        .DINT[1].4   // JY-001B Supply Pump Aux Contact
        .DINT[2].3   // JY-001A Supply Pump Enable
        .DINT[2].9   // XY-302 Chem #2 Enable
        .DINT[2].4   // XY-018 Return to Drain
        .REAL[0]   // TT-005 Supply Temperature 0-100 deg C
        .STRING[0]   // Step Name
        .STRING[1]   // Status Message
        .DINT[2].5   // AH-376 Alarm Horn
        .STRING[2]   // Step Time Remaining
        .DINT[1].0   // CP-153 Control Power On
        .STRING[3]   // Recipe Name
   Integer : DINT[150] := ([0] := 39, [1] := 39, [5] := 2, [6] := 39, [7] := 1, [8] := 7, [10] := 60, [11] := 29, [12] := 65, [15] := -2, [20] := 20, [21] := 21, [22] := 61, [26] := 120, [27] := 120, [28] := 100, [29] := 1, [36] := -4, [38] := -1, [39] := 190, [40] := 80, [41] := 80, [43] := 120, [44] := 120, [45] := 120, [46] := 120, [48] := 50, [52] := 2, [53] := -2, [54] := 2, [56] := 6242, [57] := 31208, [58] := 12, [60] := 16383, [61] := 84, [62] := 10000, [80] := 5921);   // INTEGER
        [0]   // CURRENT CIP RECIPE SELECTOR SWITCH POSITION
        [15]   // MANUAL CONTROL WORKING REGISTER
        [1]   // RECIPE SELECTOR LIST POSITION
        [30]   // MESSAGE INDEX REGISTER
        [6]   // EDIT RECIPES SELECTOR LIST POSITION
   Integer_1 : ALIAS FOR Integer[1];   // RECIPE SELECTOR LIST POSITION ALIAS
   Integer_6 : ALIAS FOR Integer[6];   // EDIT RECIPES SELECTOR LIST POSITION ALIAS
   IO_Status : INT := 16384;   // REMOTE I/O STATUS
   IO_Status_Masked : INT := 16384;   // REMOTE I/O STATUS MASK
   Message_Index : ALIAS FOR Integer[30];   // MESSAGE INDEX REGISITER
   Message_Present : INT[5];   // MESSAGES 1-80 PRESENT BITS
        [4].10   // MESSAGE 75 PRESENT
        [4].11   // MESSAGE 76 PRESENT
        [3].15   // MESSAGE 64 PRESENT
        [3].2   // MESSAGE 51 PRESENT
        [3].7   // MESSAGE 56 PRESENT
        [3].8   // MESSAGE 57 PRESENT
        [4].2   // MESSAGE 67 PRESENT
        [4].3   // MESSAGE 68 PRESENT
        [3].3   // MESSAGE 52 PRESENT
        [3].4   // MESSAGE 53 PRESENT
        [3].9   // MESSAGE 58 PRESENT
        [4]   // MESSAGES 65-80 PRESENT BITS
        [0].9   // MESSAGE 10 PRESENT
        [4].12   // MESSAGE 77 PRESENT
        [4].13   // MESSAGE 78 PRESENT
        [0].0   // MESSAGE 1 PRESENT
        [4].4   // MESSAGE 69 PRESENT
        [4].5   // MESSAGE 70 PRESENT
        [0].3   // MESSAGE 4 PRESENT
        [0].4   // MESSAGE 5 PRESENT
        [3].5   // MESSAGE 54 PRESENT
        [3].6   // MESSAGE 55 PRESENT
        [0].5   // MESSAGE 6 PRESENT
        [1].9   // MESSAGE 26 PRESENT
        [0].7   // MESSAGE 8 PRESENT
        [4].6   // MESSAGE 71 PRESENT
        [4].7   // MESSAGE 72 PRESENT
        [0]   // MESSAGES 1-16 PRESENT BITS
        [0].1   // MESSAGE 2 DEVICE IN MANUAL MODE PRESENT
        [0].10   // MESSAGE 11 PRESS "START" BUTTON TO RESUME RECIPE PRESENT
        [0].8   // MESSAGE 9 PRESENT
        [0].11   // MESSAGE 12 PRESENT
        [0].12   // MESSAGE 13 PRESENT
        [0].13   // MESSAGE 14 PRESENT
        [0].14   // MESSAGE 15 PRESENT
        [0].15   // MESSAGE 16 PRESENT
        [0].2   // MESSAGE 3 HOLD BUTTON ACTIVE PRESENT
        [0].6   // MESSAGE 7 FLOW PID CONTROLLER IN MANUAL MODE PRESENT
        [1]   // MESSAGE 17-32 PRESENT BITS
        [1].0   // MESSAGE 17 FILL HOLD PRESENT
        [1].1   // MESSAGE 18 EMPTY HOLD PRESENT
        [1].10   // MESSAGE 27 PRESENT
        [1].11   // MESSAGE 28 PRESENT
        [1].12   // MESSAGE 29 PRESENT
        [1].13   // MESSAGE 30 PRESENT
        [1].14   // MESSAGE 31 SEPARATOR TANK IN LOW LEVEL PRESENT
        [2].10   // MESSAGE 43 PRESENT
        [1].15   // MESSAGE 32 LOW LEVEL RECOVERY IN PROGRESS PRESENT
        [2]   // MESSAGES 33-48 PRESENT BITS
        [1].2   // MESSAGE 19 SUPPLY TEMPERATURE HOLD PRESENT
        [2].13   // MESSAGE 46 PRESENT
        [1].3   // MESSAGE 20 RETURN TEMPERATURE HOLD PRESENT
        [2].14   // MESSAGE 47 PRESENT
        [1].4   // MESSAGE 21 RINSE CONDUCTIVITY HOLD PRESENT
        [2].15   // MESSAGE 48 PRESENT
        [1].5   // MESSAGE 22 CHEM #1 CONDUCTIVITY HOLD PRESENT
        [2].11   // MESSAGE 44 PRESENT
        [1].6   // MESSAGE 23 CHEM #2 CONDUCTIVITY HOLD PRESENT
        [2].12   // MESSAGE 45 PRESENT
        [1].7   // MESSAGE 24 CHEM #1 INJECTION/MIX TIME HOLD PRESENT
        [2].0   // MESSAGE 33 PRESENT
        [1].8   // MESSAGE 25 CHEM #2 INJECTION/MIX TIME HOLD PRESENT
        [2].1   // MESSAGE 34 PRESENT
        [2].2   // MESSAGE 35 CHEM #1 TANK LOW LEVEL PRESENT
        [2].4   // MESSAGE 37 PRESENT
        [2].3   // MESSAGE 36 CHEM #2 TANK LOW LEVEL PRESENT
        [2].5   // MESSAGE 38 PRESENT
        [2].6   // MESSAGE 39 OVERFLOW TANK EMPTY HOLD PRESENT
        [3]   // MESSAGES 49-64 PRESENT BITS
        [2].7   // MESSAGE 40 OVERFLOW TANK HIGH LEVEL PRESENT
        [3].0   // MESSAGE 49 PRESENT
        [2].8   // MESSAGE 41 PROCESS EQUIPMENT HEARTBEAT MISSING PRESENT
        [2].9   // MESSAGE 42 PRESENT
        [3].1   // MESSAGE 50 PRESENT
        [3].10   // MESSAGE 59 PRESENT
        [4].8   // MESSAGE 73 PRESENT
        [4].9   // MESSAGE 74 PRESENT
        [4].0   // MESSAGE 65 PRESENT
        [4].1   // MESSAGE 66 PRESENT
        [4].14   // MESSAGE 79 PRESENT
        [4].15   // MESSAGE 80 PRESENT
        [3].11   // MESSAGE 60 PRESENT
        [3].12   // MESSAGE 61 PRESENT
        [3].13   // MESSAGE 62 PRESENT
        [3].14   // MESSAGE 63 PRESENT
   Message_Seq : DINT[101] := ([2] := 35, [3] := 36, [4] := 36, [5] := 36, [6] := 36, [7] := 36);   // MESSAGE SEQUENCER ARRAY
   Message_Timer : TIMER[1] := ([0].PRE := 1500, [0].ACC := 1020, [0].EN := 1, [0].TT := 1);   // MESSAGE SEQUENCER CONTROL TIMER
        [0]   // MESSAGE SCAN TIME DELAY
   Messages_List : STRING;   // ACTIVE MESSAGES ECHO FROM HMI
   MOA_Drain_Flow_Mod_Value : INT := 100;   // PV MOA DRAIN FLOW MODULATION VALUE
   MOA_Drain_Flow_Mod_Value_Ind : INT;   // PV DRAIN FLOW MODULATION VALUE STATUS
   MOA_Drain_Flow_Mod_Value_Status : BOOL;   // PV MOA DRAIN FLOW MODULATION VALUE STATUS BIT
   MOA_OFF : DINT[20];   // PANELVIEW MOA OFF
        [3]   // PV MOA SCREEN 3 MANUAL OFF BITS
        [3].0   // PV MOA SPARE MANUAL OFF
        [7].15   // PV MOA MANUAL OFF
        [7].2   // PV MOA MANUAL OFF
        [4].10   // PV MOA SPARE MANUAL OFF
        [4].11   // PV MOA SPARE MANUAL OFF
        [1].13   // PV MOA CHEM #2 BLOCK XY-305 MANUAL OFF
        [5].1   // PV MOA MANUAL OFF
        [5].3   // PV MOA MANUAL OFF
        [5].4   // PV MOA MANUAL OFF
        [1].5   // PV MOA RETURN TO DRAIN XY-018 MANUAL OFF
        [3].16   // PV MOA MANUAL OFF
        [3].3   // PV MOA SPARE MANUAL OFF
        [3].4   // PV MOA SPARE MANUAL OFF
        [5].5   // PV MOA MANUAL OFF
        [5].6   // PV MOA MANUAL OFF
        [1].6   // PV MOA ALARM HORN AH-376 MANUAL OFF
        [2].10   // PV MOA SPARE MANUAL OFF
        [3].5   // PV MOA SPARE MANUAL OFF
        [3].6   // PV MOA SPARE MANUAL OFF
        [5].7   // PV MOA MANUAL OFF
        [5].8   // PV MOA MANUAL OFF
        [1].7   // PV MOA HEATER ENABLE JY-004A MANUAL OFF
        [5].12   // PV MOA MANUAL OFF
        [7].13   // PV MOA MANUAL OFF
        [7].14   // PV MOA MANUAL OFF
        [1].14   // PV MOA OVERFLOW TANK DRAIN PUMP XV-032 MANUAL OFF
        [6].13   // PV MOA MANUAL OFF
        [6].14   // PV MOA MANUAL OFF
        [1]   // PV MOA SCREEN 1 MANUAL OFF BITS
        [1].0   // PV MOA SPARE OUT-396 MANUAL OFF
        [6].3   // PV MOA MANUAL OFF
        [6].4   // PV MOA MANUAL OFF
        [6].5   // PV MOA MANUAL OFF
        [6].6   // PV MOA MANUAL OFF
        [7].5   // PV MOA MANUAL OFF
        [7].6   // PV MOA MANUAL OFF
        [1].15   // PV MOA SPARE OUT-396 MANUAL OFF
        [2].12   // PV MOA SPARE MANUAL OFF
        [6].7   // PV MOA MANUAL OFF
        [6].8   // PV MOA MANUAL OFF
        [6].9   // PV MOA MANUAL OFF
        [7].0   // PV MOA MANUAL OFF
        [7].7   // PV MOA MANUAL OFF
        [7].8   // PV MOA MANUAL OFF
        [1].16   // PV MOA DRAIN FLOW MODULATION VALVE MANUAL OFF
        [1].1   // PV MOA AIR BLOW XV-008A MANUAL OFF
        [2].11   // PV MOA SPARE MANUAL OFF
        [3].7   // PV MOA SPARE MANUAL OFF
        [3].8   // PV MOA SPARE MANUAL OFF
        [3].1   // PV MOA SPARE MANUAL OFF
        [3].10   // PV MOA SPARE MANUAL OFF
        [3].11   // PV MOA SPARE MANUAL OFF
        [3].12   // PV MOA SPARE MANUAL OFF
        [1].8   // PV MOA AIR BLOW BLOCK XY-008 MANUAL OFF
        [5].13   // PV MOA MANUAL OFF
        [1].2   // PV MOA SUPPLY PUMP CASING DRAIN XY-002 MANUAL OFF
        [1].9   // PV MOA SPARE OUT-384 MANUAL OFF
        [2]   // PV MOA SCREEN 2 MANUAL OFF BITS
        [7].1   // PV MOA MANUAL OFF
        [7].10   // PV MOA MANUAL OFF
        [1].10   // PV MOA CHEM #1 ENABLE XY-202 MANUAL OFF
        [5].9   // PV MOA MANUAL OFF
        [6].0   // PV MOA MANUAL OFF
        [2].13   // PV MOA SPARE MANUAL OFF
        [2].14   // PV MOA SPARE MANUAL OFF
        [7].9   // PV MOA MANUAL OFF
        [2].15   // PV MOA SPARE MANUAL OFF
        [2].5   // PV MOA SPARE OUT-414 MANUAL OFF
        [6].1   // PV MOA MANUAL OFF
        [6].10   // PV MOA MANUAL OFF
        [2].2   // PV MOA DRAIN TO WASTE NEUTRALIZATION XY-024 MANUAL OFF
        [4].2   // PV MOA SPARE MANUAL OFF
        [4].3   // PV MOA SPARE MANUAL OFF
        [7].11   // PV MOA MANUAL OFF
        [7].12   // PV MOA MANUAL OFF
        [4].12   // PV MOA SPARE MANUAL OFF
        [4].13   // PV MOA SPARE MANUAL OFF
        [3].9   // PV MOA SPARE MANUAL OFF
        [4]   // PV MOA SCREEN 4 MANUAL OFF BITS
        [3].13   // PV MOA SPARE MANUAL OFF
        [3].14   // PV MOA SPARE MANUAL OFF
        [4].4   // PV MOA SPARE MANUAL OFF
        [4].5   // PV MOA SPARE MANUAL OFF
        [2].0   // PV MOA OVERFLOW TANK DRAIN XY-022 MANUAL OFF
        [2].3   // PV MOA SPARE SOLENOID SV-410 MANUAL OFF
        [5].14   // PV MOA MANUAL OFF
        [4].6   // PV MOA SPARE MANUAL OFF
        [4].7   // PV MOA SPARE MANUAL OFF
        [1].11   // PV MOA CHEM #2 ENABLE XY-302 MANUAL OFF
        [4].8   // PV MOA SPARE MANUAL OFF
        [4].9   // PV MOA SPARE MANUAL OFF
        [6].15   // PV MOA MANUAL OFF
        [6].2   // PV MOA MANUAL OFF
        [5]   // PV MOA SCREEN 5 MANUAL OFF BITS
        [5].2   // PV MOA MANUAL OFF
        [2].4   // PV MOA SPARE SOLENOID SV-412 MANUAL OFF
        [5].15   // PV MOA MANUAL OFF
        [1].12   // PV MOA CHEM #1 BLOCK XY-205 MANUAL OFF
        [5].0   // PV MOA MANUAL OFF
        [6].11   // PV MOA MANUAL OFF
        [6].12   // PV MOA MANUAL OFF
        [2].6   // PV MOA SPARE OUT-416 MANUAL OFF
        [2].8   // PV MOA SPARE MANUAL OFF
        [2].7   // PV MOA SPARE OUT-418 MANUAL OFF
        [2].9   // PV MOA SPARE MANUAL OFF
        [3].15   // PV MOA SPARE MANUAL OFF
        [3].2   // PV MOA SPARE MANUAL OFF
        [1].3   // PV MOA SUPPLY PUMP ENABLE JY-001A MANUAL OFF
        [1].4   // PV MOA SPARE SOLENOID SV-372 MANUAL OFF
        [5].10   // PV MOA MANUAL OFF
        [7].3   // PV MOA MANUAL OFF
        [7].4   // PV MOA MANUAL OFF
        [4].14   // PV MOA SPARE MANUAL OFF
        [4].15   // PV MOA SPARE MANUAL OFF
        [4].0   // PV MOA SPARE MANUAL OFF
        [4].1   // PV MOA SPARE MANUAL OFF
        [2].1   // PV MOA LOW POINT DRAIN XY-023 MANUAL OFF
        [5].11   // PV MOA MANUAL OFF
   MOA_ON : DINT[20];   // PANELVIEW MOA ON
        [6].12   // PV MOA MANUAL ON
        [6].13   // PV MOA MANUAL ON
        [6].14   // PV MOA MANUAL ON
        [6].15   // PV MOA MANUAL ON
        [6].5   // PV MOA MANUAL ON
        [6].6   // PV MOA MANUAL ON
        [6].7   // PV MOA MANUAL ON
        [6].8   // PV MOA MANUAL ON
        [6].9   // PV MOA MANUAL ON
        [7]   // PV MOA SCREEN 7 MANUAL ON BITS
        [3].2   // PV MOA SPARE MANUAL ON
        [3].3   // PV MOA SPARE MANUAL ON
        [5].6   // PV MOA MANUAL ON
        [7].0   // PV MOA MANUAL ON
        [7].1   // PV MOA MANUAL ON
        [3].4   // PV MOA SPARE MANUAL ON
        [3].5   // PV MOA SPARE MANUAL ON
        [4].11   // PV MOA SPARE MANUAL ON
        [4].12   // PV MOA SPARE MANUAL ON
        [5].7   // PV MOA MANUAL ON
        [7].8   // PV MOA MANUAL ON
        [7].9   // PV MOA MANUAL ON
        [5].8   // PV MOA MANUAL ON
        [4].13   // PV MOA SPARE MANUAL ON
        [4].14   // PV MOA SPARE MANUAL ON
        [3].6   // PV MOA SPARE MANUAL ON
        [3].7   // PV MOA SPARE MANUAL ON
        [5].9   // PV MOA MANUAL ON
        [6].0   // PV MOA MANUAL ON
        [4].15   // PV MOA SPARE MANUAL ON
        [4].2   // PV MOA SPARE MANUAL ON
        [5].0   // PV MOA MANUAL ON
        [6].1   // PV MOA MANUAL ON
        [4].3   // PV MOA SPARE MANUAL ON
        [4].4   // PV MOA SPARE MANUAL ON
        [7].10   // PV MOA MANUAL ON
        [7].11   // PV MOA MANUAL ON
        [3].8   // PV MOA SPARE MANUAL ON
        [3].9   // PV MOA SPARE MANUAL ON
        [4].5   // PV MOA SPARE MANUAL ON
        [4].6   // PV MOA SPARE MANUAL ON
        [7].12   // PV MOA MANUAL ON
        [7].13   // PV MOA MANUAL ON
        [1]   // PV MOA SCREEN 1 MANUAL ON BITS
        [7].14   // PV MOA MANUAL ON
        [7].15   // PV MOA MANUAL ON
        [5].1   // PV MOA MANUAL ON
        [6].2   // PV MOA MANUAL ON
        [4]   // PV MOA SCREEN 4 MANUAL ON BITS
        [4].0   // PV MOA SPARE MANUAL ON
        [6].3   // PV MOA MANUAL ON
        [5].10   // PV MOA MANUAL ON
        [5].11   // PV MOA MANUAL ON
        [7].2   // PV MOA MANUAL ON
        [7].3   // PV MOA MANUAL ON
        [4].7   // PV MOA SPARE MANUAL ON
        [4].8   // PV MOA SPARE MANUAL ON
        [2].9   // PV MOA SPARE MANUAL ON
        [5].2   // PV MOA MANUAL ON
        [6].4   // PV MOA MANUAL ON
        [1].0   // PV MOA SPARE OUT-396 MANUAL ON
        [2].10   // PV MOA SPARE MANUAL ON
        [5].3   // PV MOA MANUAL ON
        [4].1   // PV MOA SPARE MANUAL ON
        [4].10   // PV MOA SPARE MANUAL ON
        [1].1   // PV MOA AIR BLOW XV-008A MANUAL ON
        [5].14   // PV MOA MANUAL ON
        [1].10   // PV MOA CHEM #1 ENABLE XY-202 MANUAL ON
        [1].11   // PV MOA CHEM #2 ENABLE XY-302 MANUAL ON
        [1].12   // PV MOA CHEM #1 BLOCK XY-205 MANUAL ON
        [1].13   // PV MOA CHEM #2 BLOCK XY-305 MANUAL ON
        [1].14   // PV MOA OVERFLOW TANK DRAIN PUMP XV-032 MANUAL ON
        [1].15   // PV MOA SPARE OUT-396 MANUAL ON
        [2].8   // PV MOA SPARE MANUAL ON
        [1].16   // PV MOA DRAIN FLOW MODULATION VALVE MANUAL ON
        [1].2   // PV MOA SUPPLY PUMP CASING DRAIN XY-002 MANUAL ON
        [1].3   // PV MOA SUPPLY PUMP ENABLE JY-001A MANUAL ON
        [1].4   // PV MOA SPARE SOLENOID SV-372 MANUAL ON
        [1].5   // PV MOA RETURN TO DRAIN XY-018 MANUAL ON
        [1].6   // PV MOA ALARM HORN AH-376 MANUAL ON
        [5].12   // PV MOA MANUAL ON
        [1].7   // PV MOA HEATER ENABLE JY-004A MANUAL ON
        [1].8   // PV MOA AIR BLOW BLOCK XY-008 MANUAL ON
        [1].9   // PV MOA SPARE OUT-384 MANUAL ON
        [2].11   // PV MOA SPARE MANUAL ON
        [2]   // PV MOA SCREEN 2 MANUAL ON BITS
        [2].12   // PV MOA SPARE MANUAL ON
        [2].0   // PV MOA OVERFLOW TANK DRAIN XY-022 MANUAL ON
        [2].1   // PV MOA LOW POINT DRAIN XY-023 MANUAL ON
        [2].13   // PV MOA SPARE MANUAL ON
        [2].14   // PV MOA SPARE MANUAL ON
        [2].15   // PV MOA SPARE MANUAL ON
        [2].5   // PV MOA SPARE OUT-414 MANUAL ON
        [2].2   // PV MOA DRAIN TO WASTE NEUTRALIZATION XY-024 MANUAL ON
        [2].3   // PV MOA SPARE SOLENOID SV-410 MANUAL ON
        [2].4   // PV MOA SPARE SOLENOID SV-412 MANUAL ON
        [5].4   // PV MOA MANUAL ON
        [5].13   // PV MOA MANUAL ON
        [2].6   // PV MOA SPARE OUT-416 MANUAL ON
        [3].1   // PV MOA SPARE MANUAL ON
        [4].9   // PV MOA SPARE MANUAL ON
        [5]   // PV MOA SCREEN 5 MANUAL ON BITS
        [7].4   // PV MOA MANUAL ON
        [7].5   // PV MOA MANUAL ON
        [5].5   // PV MOA MANUAL ON
        [2].7   // PV MOA SPARE OUT-418 MANUAL ON
        [3].10   // PV MOA SPARE MANUAL ON
        [7].6   // PV MOA MANUAL ON
        [7].7   // PV MOA MANUAL ON
        [3]   // PV MOA SCREEN 3 MANUAL ON BITS
        [3].11   // PV MOA SPARE MANUAL ON
        [5].15   // PV MOA MANUAL ON
        [6]   // PV MOA SCREEN 6 MANUAL ON BITS
        [3].0   // PV MOA SPARE MANUAL ON
        [3].12   // PV MOA SPARE MANUAL ON
        [3].13   // PV MOA SPARE MANUAL ON
        [3].14   // PV MOA SPARE MANUAL ON
        [3].15   // PV MOA SPARE MANUAL ON
        [6].10   // PV MOA MANUAL ON
        [6].11   // PV MOA MANUAL ON
   MOA_One_Shot : BOOL[32];   // PANELVIEW MOA ONE SHOT
   MOA_Screen1_Auto : BOOL;   // PV MOA SCREEN #1 AUTO PB
   MOA_Screen1_Man_Off : BOOL;   // PV MOA SCREEN #1 OFF PB
   MOA_Screen1_Man_On : BOOL;   // PV MOA SCREEN #1 MANUAL PB
   MOA_Screen2_Auto : BOOL;   // PV MOA SCREEN #2 AUTO PB
   MOA_Screen2_Man_Off : BOOL;   // PV MOA SCREEN #2 OFF PB
   MOA_Screen2_Man_On : BOOL;   // PV MOA SCREEN #2 MANUAL PB
   MOA_Select : DINT[10] := ([1] := 1, [2] := 2, [3] := 1, [4] := 64, [5] := 128, [6] := 1);   // MAN/OFF/AUTO SELECT
        [1]   // MOA SELECT SCREEN 1
        [3]   // MOA SELECT SCREEN 3
        [4]   // MOA SELECT SCREEN 4
        [5]   // MOA SELECT SCREEN 5
        [6]   // MOA SELECT SCREEN 6
        [7]   // MOA SELECT SCREEN 7
        [8]   // MOA SELECT SCREEN 8
        [9]   // MOA SELECT SCREEN 9
        [2]   // MOA SELECT SCREEN 2
   MOA_Status : DINT[10];   // MAN/OFF/AUTO STATUS
        [1]   // MOA SCREEN 1 STATUS
        [2]   // MOA SCREEN 2 STATUS
        [3]   // MOA SCREEN 3 STATUS
        [4]   // MOA SCREEN 4 STATUS
        [5]   // MOA SCREEN 5 STATUS
        [6]   // MOA SCREEN 6 STATUS
        [7]   // MOA SCREEN 7 STATUS
        [8]   // MOA SCREEN 8 STATUS
        [9]   // MOA SCREEN 9 STATUS
   One_Shot : BOOL[128] := ([10] := 1, [11] := 1, [12] := 1, [13] := 1, [14] := 1, [15] := 1, [16] := 1, [17] := 1, [29] := 1, [30] := 1, [31] := 1, [32] := 1, [39] := 1);   // ONE SHOT ARRAY
        [10]   // ONE SHOT
        [11]   // ONE SHOT
        [1]   // ONE SHOT
        [12]   // ONE SHOT
        [3]   // ONE SHOT
        [13]   // ONE SHOT
        [14]   // ONE SHOT
        [15]   // ONE SHOT
        [16]   // ONE SHOT
        [17]   // ONE SHOT
        [36]   // PANELVIEW RTC HOURLY UPDATE SIGNAL FROM PLC HOURLY CLOCK UPDATE ONE-SHOT
        [39]   // ONE SHOT
        [40]   // ONE SHOT
        [74]   // ONE SHOT
        [5]   // ONE SHOT
        [37]   // PANELVIEW RTC HOURLY UPDATE SIGNAL FROM HMI CLOCK UPDATE ONE-SHOT
        [7]   // ONE SHOT
        [8]   // ONE SHOT
        [9]   // ONE SHOT
   Opcode_Description : STRING;   // ACTIVE OPCODE ECHO FROM HMI
   OpCode_Pin : DINT[5];   // OPCODE PIN ARRAY
        [1].9   // SEQ PIN WORD #1 PIN #09 EMPTY HOLD
        [4].13   // SEQ PIN WORD #4 PIN #13
        [4].4   // SEQ PIN WORD #4 PIN #04
        [3].15   // SEQ PIN WORD #3 PIN #15
        [3].6   // SEQ PIN WORD #3 PIN #06
        [2].4   // SEQ PIN WORD #2 PIN #04 PRE-HEAT
        [2].5   // SEQ PIN WORD #2 PIN #05
        [2].6   // SEQ PIN WORD #2 PIN #06
        [4].14   // SEQ PIN WORD #4 PIN #14
        [4].5   // SEQ PIN WORD #4 PIN #05
        [1]   // SEQUENCER OUTPUTS WORD #1
        [3].10   // SEQ PIN WORD #3 PIN #10
        [3].2   // SEQ PIN WORD #3 PIN #02
        [4].15   // SEQ PIN WORD #4 PIN #15
        [4].6   // SEQ PIN WORD #4 PIN #06
        [3].11   // SEQ PIN WORD #3 PIN #11
        [3].3   // SEQ PIN WORD #3 PIN #03
        [4].7   // SEQ PIN WORD #4 PIN #07
        [4].8   // SEQ PIN WORD #4 PIN #08
        [3].12   // SEQ PIN WORD #3 PIN #12
        [3].4   // SEQ PIN WORD #3 PIN #04
        [1].0   // SEQ PIN WORD #1 PIN #00 AWFI FILL ON
        [2].10   // SEQ PIN WORD #2 PIN #10 TEMP 2 ( RINSE)
        [3].13   // SEQ PIN WORD #3 PIN #13
        [3].5   // SEQ PIN WORD #3 PIN #05
        [3].8   // SEQ PIN WORD #3 PIN #08
        [4].0   // SEQ PIN WORD #4 PIN #00
        [2].7   // SEQ PIN WORD #2 PIN #07 TEMP 5 (FINAL RINSE)
        [1].1   // SEQ PIN WORD #1 PIN #01
        [3]   // SEQUENCER OUTPUTS WORD #3
        [2].11   // SEQ PIN WORD #2 PIN #11 TEMP 1 (PRE-RINSE)
        [1].14   // SEQ PIN WORD #1 PIN #14
        [2]   // SEQUENCER OUTPUTS WORD #2
        [1].15   // SEQ PIN WORD #1 PIN #15 LOW LEVEL DISABLE
        [2].8   // SEQ PIN WORD #2 PIN #08 TEMP 4 (CHEM #2 WASH)
        [1].2   // SEQ PIN WORD #1 PIN #02 LOW POINT DRAIN
        [4].1   // SEQ PIN WORD #4 PIN #01
        [4].10   // SEQ PIN WORD #4 PIN #10
        [4].9   // SEQ PIN WORD #4 PIN #09
        [2].12   // SEQ PIN WORD #2 PIN #12
        [4]   // SEQUENCER OUTPUTS WORD #4
        [2].9   // SEQ PIN WORD #2 PIN #09 TEMP 3 (CHEM #1 WASH)
        [1].10   // SEQ PIN WORD #1 PIN #10 RINSE CONDUCTIVITY HOLD
        [4].11   // SEQ PIN WORD #4 PIN #11
        [4].2   // SEQ PIN WORD #4 PIN #02
        [1].3   // SEQ PIN WORD #1 PIN #03 PAUSE
        [2].0   // SEQ PIN WORD #2 PIN #00 CHEM #2 CONDUCTIVITY
        [2].13   // SEQ PIN WORD #2 PIN #13 FLOW CONTROL ENABLE
        [3].1   // SEQ PIN WORD #3 PIN #01
        [3].7   // SEQ PIN WORD #3 PIN #07
        [3].14   // SEQ PIN WORD #3 PIN #14
        [3].9   // SEQ PIN WORD #3 PIN #09
        [2].14   // SEQ PIN WORD #2 PIN #14
        [2].15   // SEQ PIN WORD #2 PIN #15 SUPPLY PUMP
        [4].12   // SEQ PIN WORD #4 PIN #12
        [4].3   // SEQ PIN WORD #4 PIN #03
        [1].4   // SEQ PIN WORD #1 PIN #04 MODULATION DRAIN VALVE
        [1].5   // SEQ PIN WORD #1 PIN #05 PUMP CASING DRAIN
        [2].2   // SEQ PIN WORD #2 PIN #02 OVERFLOW TANK DRAIN PUMP
        [2].3   // SEQ PIN WORD #2 PIN #03
        [3].0   // SEQ PIN WORD #3 PIN #00
        [1].6   // SEQ PIN WORD #1 PIN #06 RETURN LINE DRAIN
        [1].7   // SEQ PIN WORD #1 PIN #07 AIR BLOW
        [1].11   // SEQ PIN WORD #1 PIN #11 WASH CONDUCTIVITY HOLD
        [1].12   // SEQ PIN WORD #1 PIN #12 TEMPERATURE HOLD
        [2].1   // SEQ PIN WORD #2 PIN #01 CHEM #1 CONDUCTIVITY
        [1].8   // SEQ PIN WORD #1 PIN #08
        [1].13   // SEQ PIN WORD #1 PIN #13 FILL HOLD
   OpCode_Word : DINT[5,97] := ([1,2] := 16#0000_8274, [1,4] := 16#0000_a001, [1,5] := 16#0000_8214, [1,7] := 16#0000_1000, [1,8] := 16#0000_1001, [1,9] := 16#0000_0015, [1,10] := 16#0000_1801, [1,11] := 16#0000_1801, [1,13] := 16#0000_1001, [1,14] := 16#0000_0415, [1,16] := 16#0000_0015, [1,17] := 16#0000_0095, [1,18] := 16#0000_0200, [1,20] := 16#0000_0008, [2,2] := 16#0000_2000, [2,5] := 16#0000_8000, [2,7] := 16#0000_8010, [2,8] := 16#0000_a800, [2,9] := 16#0000_a800, [2,10] := 16#0000_a202, [2,11] := 16#0000_a101, [2,13] := 16#0000_a400, [2,14] := 16#0000_a080, [2,16] := 16#0000_a400, [2,17] := 16#0000_8000, [2,18] := 16#0000_0004);   // OPCODE WORD ARRAY
        [1,0]   // OPCODE WORD #1
        [2,0]   // OPCODE WORD #2
        [3,0]   // OPCODE WORD #3
        [4,0]   // OPCODE WORD #4
   Panelview : INT[40] := ([0] := 2048, [4] := 20, [6] := 1, [7] := 1, [14] := 1, [15] := 1, [20] := 2, [31] := 1, [32] := 1, [33] := 75, [34] := -1);   // PANELVIEW CONTROL
        [8].0   // CYCLE SELECT
        [31]   // PANELVIEW TERMINAL CURRENT DISPLAY STATUS
        [4]   // TOTAL NUMBER OF STEPS IN RECIPE
        [0]   // PANELVIEW PUSHBUTTON
        [0].0   // PANELVIEW START
        [0].1   // PANELVIEW STOP
        [0].2   // PANELVIEW HOLD
        [0].7   // PANELVIEW MANUAL STEP
        [0].3   // PANELVIEW ABORT
        [0].5   // PANELVIEW UPDATE CLOCK PUSHBUTTON
        [0].6   // PANELVIEW PRINT
        [0].15   // ALL OUTPUTS TO AUTO
        [16].0   // PANELVIEW RECIPE RENAME NOTIFICATION
        [16].1   // PANELVIEW RECIPE RENAME HANDSHAKE
        [21]   // PANELVIEW TERMINAL CONTROL
        [2]   // PANELVIEW RTC HOURLY UPDATE
   PID2 : PID := (CTL := -2080340224, EN := 1, SWM := 1, INI := 1, DVNA := 1, DVPA := 1, PVLA := 1, KP := 0.5, KI := 0.1, BIAS := -0.030520372, MAXS := 60.0, DB := 1.0, MAXO := 100.0, UPD := 0.25, PVH := 16383.0, MAXI := 60.0, MAXCV := 16383.0, MAXTIE := 60.0, DATA[0] := 0.030520372, DATA[5] := 1.6666666, DATA[6] := 1.0, DATA[7] := 4.0, DATA[8] := 0.5, DATA[9] := 0.1, DATA[11] := 0.5, DATA[12] := 0.1, DATA[15] := 163.83, DATA[16] := 1.6666666);   // SUPPLY FLOW PID
   PID2_bumpless_transfer : BOOL;   // FORCE PID TO RESTART FROM PREVIOUS OUTPUT VALUE
   PID2_Man_Mode : BOOL;   // PID2 MANUAL MODE
   PID2_Manual_PB_Pressed : BOOL;   // PID2 MANUAL PUSHBUTTON PRESSED
   PID2_Output_Memory : REAL;   // SUPPLY FLOW PID OUTPUT MEMORY TO USE FOR BUMPLESS TRANSFER
   PID2_PV_Manual_PB : BOOL;   // PID2 MANUAL MODE SELECTED ON HMI
   PID2_Setpoint_Memory : REAL := 35.0;   // SUPPLY FLOW PID SETPOINT MEMORY TO USE FOR BUMPLESS TRANSFER
   PID_Ons : DINT[6] := ([2] := 966, [5] := 1014);   // PID ONE SHOT
        [0].0   // ONE SHOT
        [0].1   // ONE SHOT
        [0].2   // ONE SHOT
        [0].3   // ONE SHOT
        [2].0   // PID 2 ONE SHOT
        [3].1   // PID 3 ONE SHOT
        [2].1   // PID 2 ONE SHOT
        [2].2   // PID 2 ONE SHOT
        [2].3   // PID 2 ONE SHOT
        [2].4   // PID 2 ONE SHOT
        [4].1   // PID 4 ONE SHOT
        [2].6   // PID 2 ONE SHOT
        [5].1   // PID 5 ONE SHOT
   PID_Timer : TIMER[5] := ([0].PRE := 5000, [0].ACC := 5000, [0].EN := 1, [0].DN := 1, [1].PRE := 8000, [2].PRE := 5000, [2].EN := 1, [2].DN := 1, [3].PRE := 8000, [4].PRE := 50, [4].ACC := 51, [4].EN := 1, [4].DN := 1);   // PID TIMERS
        [2]   // PID2 OUTPUT IS FORCED TO ZERO FOR A PRESET AMOUNT OF TIME.
        [3]   // PID 2 DELAY START OF AUTO MODE TO ALLOW FLOW TO PICK UP WHERE IT LEFT OFF
        [4]   // PID 2 DELAY UNLATCH OF MANUAL MODE TO ALLOW THE PID2.SO TO GO TO ZERO BEFORE UNLATCHING THE MANUAL MODE
   Process_Heartbeat_Memory : BOOL;
   Process_to_CIP : Process_to_CIP;   // PROCESS SIGNALS TO CIP
        .DINT[0].0   // Heartbeat Signal from DCS
        .DINT[0].1   // DCS Remote Process Stop
        .REAL[0]   // CIP Remote Flow Setpoint 0-60 GPM
   PV_Copy_Recipes_Destination : DINT := 35;   // COPY RECIPES DESTINATION
   PV_Copy_Recipes_Duration : TIMER := (PRE := 1000);   // COPY RECIPES COPY DURATION
   PV_Copy_Recipes_One_Shot : BOOL;   // COPY RECIPES REQUEST TO COPY ONE SHOT
   PV_Copy_Recipes_Request : BOOL;   // COPY RECIPES REQUEST TO COPY
   PV_Copy_Recipes_Source : DINT := 34;
   PV_Current_Select_Step_Op : DINT;   // PANELVIEW STORES CURRENT OPCODE NUMBER OF STEP BEING EDITED FOR DISPLAY ON OPCODE LIST SCREEN
   PV_Edit_OpCode_List : DINT[24] := ([1] := 1, [2] := 2, [3] := 3, [4] := 4, [5] := 5, [6] := 6, [7] := 7, [8] := 8, [9] := 9, [10] := 10, [11] := 11, [12] := 12, [13] := 13, [14] := 14, [15] := 15, [16] := 16, [17] := 17, [18] := 18, [19] := 19, [20] := 20, [21] := 21, [22] := 22);   // PANELVIEW RECIPE EDIT OPCODE LIST
   PV_Edit_Opcode_Sel_Top_Row : DINT := 1;   // PANELVIEW RECIPE EDIT OPCODE LIST TOP ROW #
   PV_Edit_Opcodes : DINT[300] := ([1] := 4, [2] := 8, [3] := 9, [4] := 5, [5] := 4, [6] := 7, [7] := 10, [8] := 13, [9] := 16, [10] := 20, [11] := 5, [12] := 4, [13] := 11, [14] := 13, [15] := 16, [16] := 14, [17] := 17, [18] := 18, [19] := 2, [20] := 1);   // PANELVIEW BUFFER TO EDIT OPCODES
        [0]   // EDIT RECIPES TEMPLATE OPCODE FILE
   PV_Edit_Recipe_Name : STRING := 'FAT TEST RECIPE';   // SELECTED RECIPE TO EDIT
   PV_Edit_Recipe_Top_Row : DINT := 6;   // PANELVIEW RECIPE EDIT TOP ROW #
   PV_Edit_Recipes : DINT[7] := ([0] := 26, [2] := 601);   // PANELVIEW RECIPE EDITING
        [0]   // EDIT RECIPES STEP #
        [5].3   // PV EDIT RECIPES NEW TIME HANDSHAKE
        [3].2   // EDIT RECIPES REQUEST TO SAVE
        [5].4   // PV EDIT RECIPES SELECT NEW OPCODE FROM OPCODE LIST NOTIFICATION
        [2]   // EDIT RECIPES TIME
        [5].6   // PV EDIT RECIPES NEW MINUTES NOTIFICATION
        [3].3   // EDIT RECIPES RETURN TO STEP #1
        [5].7   // PV EDIT RECIPES NEW MINUTES HANDSHAKE
        [5].0   // PV EDIT RECIPES NEW OPCODE NOTIFICATION
        [5].1   // PV EDIT RECIPES NEW OPCODE HANDSHAKE
        [5].12   // PV EDIT RECIPES NEW SECONDS NOTIFICATION
        [5].13   // PV EDIT RECIPES NEW SECONDS HANDSHAKE
        [5].2   // PV EDIT RECIPES NEW TIME NOTIFICATION
        [3].0   // PANELVIEW RECIPE EDIT SCREEN INSERT BUTTON
        [1]   // EDIT RECIPES OPCODE
        [3].1   // PANELVIEW RECIPE EDIT SCREEN DELETE BUTTON
   PV_Edit_Recipes_0 : ALIAS FOR PV_Edit_Recipes[0];   // EDIT RECIPES STEP NUMBER
   PV_Edit_Recipes_0_Prev : DINT;   // EDIT RECIPE STEP NUMBER PREVIOUS POSITION
   PV_Edit_Screen_Opcodes : DINT[25] := ([1] := 7, [2] := 10, [3] := 13, [4] := 16, [5] := 20, [6] := 5, [7] := 4, [8] := 11, [9] := 13, [10] := 16, [11] := 14, [12] := 17, [13] := 18, [14] := 2, [15] := 1);   // PANELVIEW RECIPE EDIT DISPLAY OPCODES
        [12]   // EDIT RECIPES OPCODE TEXT ROW #12
        [6]   // EDIT RECIPES OPCODE TEXT ROW #6
        [13]   // EDIT RECIPES OPCODE TEXT ROW #13
        [7]   // EDIT RECIPES OPCODE TEXT ROW #7
        [14]   // EDIT RECIPES OPCODE TEXT ROW #14
        [15]   // EDIT RECIPES OPCODE TEXT ROW #15
        [16]   // EDIT RECIPES OPCODE TEXT ROW #16
        [1]   // EDIT RECIPES OPCODE TEXT ROW #1
        [8]   // EDIT RECIPES OPCODE TEXT ROW #8
        [9]   // EDIT RECIPES OPCODE TEXT ROW #9
        [2]   // EDIT RECIPES OPCODE TEXT ROW #2
        [3]   // EDIT RECIPES OPCODE TEXT ROW #3
        [4]   // EDIT RECIPES OPCODE TEXT ROW #4
        [5]   // EDIT RECIPES OPCODE TEXT ROW #5
        [10]   // EDIT RECIPES OPCODE TEXT ROW #10
        [11]   // EDIT RECIPES OPCODE TEXT ROW #11
   PV_Edit_Setpoints : REAL[97] := ([1] := 55.0, [2] := 65.0, [3] := 60.0, [4] := 45.0, [5] := 65.0, [7] := 53.0, [8] := 63.0, [9] := 57.0, [10] := 43.0, [11] := 63.0, [13] := 85.0, [14] := 300.0, [15] := 900.0, [17] := 15.0, [18] := 14.0, [19] := 15.0, [20] := 45.0, [21] := 5.0, [22] := 15.0, [23] := 300.0, [25] := 10.0, [26] := 9.0, [27] := 10.0, [28] := 50.0, [29] := 3.0, [30] := 17.0, [31] := 300.0, [33] := 2.0, [34] := 900.0, [37] := 35.0, [41] := 5.0, [42] := 50.0, [43] := 5.0, [44] := 60.0, [45] := 50.0, [47] := 15.0, [49] := 180.0, [50] := 180.0, [52] := 30.0, [53] := 5.0, [54] := 5.0, [55] := 3.0, [57] := 300.0);   // PANELVIEW BUFFER TO EDIT SETPOINTS
        [0]   // EDIT RECIPES TEMPLATE SETPOINT FILE
   PV_Edit_Times : DINT[300] := ([1] := 10, [2] := 10, [3] := 10, [4] := 10, [5] := 10, [6] := 10, [7] := 10, [8] := 10, [9] := 10, [10] := 10, [11] := 10, [12] := 10, [13] := 10, [14] := 10, [15] := 10, [16] := 10, [17] := 10, [18] := 10, [19] := 10, [20] := 10);   // PANELVIEW BUFFER TO EDIT STEP TIMES
        [0]   // EDIT RECIPES TEMPLATE TIME FILE
   PV_Edit_Times_Indexer : DINT := 12;
   PV_Edit_Times_Minutes : DINT[98];
   PV_Edit_Times_Seconds : DINT[98] := ([1] := 10, [2] := 10, [3] := 10, [4] := 10, [5] := 10, [6] := 10, [7] := 10, [8] := 10, [9] := 10, [10] := 10, [11] := 10, [12] := 10, [13] := 10, [14] := 10, [15] := 10, [16] := 10, [17] := 10, [18] := 10, [19] := 10, [20] := 10);
   PV_Message : DINT[3] := ([2] := 5);   // PANELVIEW STATUS MESSAGE
        [0]   // MESSAGE SEQ OUTPUT WORD
        [2]   // PANELVIEW MESSAGE BUFFER
        [1]   // PANELVIEW CIP CONTROL MESSAGE
   PV_Output_Status : INT[20] := ([1] := 64);   // PV OUTPUT STATUS:
        [3].15   // PV OUTPUT STATUS: SPARE
        [4].4   // PV OUTPUT STATUS: SPARE
        [8]   // PV OUTPUT STATUS: SCREEN 8
        [3].2   // PV OUTPUT STATUS: SPARE
        [0]   // PV OUTPUT STATUS: NOT USED
        [9]   // PV OUTPUT STATUS: SCREEN 9
        [4].10   // PV OUTPUT STATUS: SPARE
        [4].5   // PV OUTPUT STATUS: SPARE
        [2].1   // PV OUTPUT STATUS: LOW POINT DRAIN XY-023
        [3].3   // PV OUTPUT STATUS: SPARE
        [1].14   // PV OUTPUT STATUS: OVERFLOW TANK DRAIN PUMP XV-032
        [4].6   // PV OUTPUT STATUS: SPARE
        [4].7   // PV OUTPUT STATUS: SPARE
        [1].15   // PV OUTPUT STATUS: SPARE OUT-396
        [4].8   // PV OUTPUT STATUS: SPARE
        [4].11   // PV OUTPUT STATUS: SPARE
        [1]   // PV OUTPUT STATUS: SCREEN 1
        [2].10   // PV OUTPUT STATUS: SPARE
        [2].11   // PV OUTPUT STATUS: SPARE
        [1].2   // PV OUTPUT STATUS: SUPPLY PUMP CASING DRAIN XY-002
        [2].12   // PV OUTPUT STATUS: SPARE
        [2].13   // PV OUTPUT STATUS: SPARE
        [1].3   // PV OUTPUT STATUS: SUPPLY PUMP ENABLE JY-001A
        [1].0   // PV OUTPUT STATUS: SPARE OUT-396
        [3]   // PV OUTPUT STATUS: SCREEN 3
        [2].14   // PV OUTPUT STATUS: SPARE
        [2].15   // PV OUTPUT STATUS: SPARE
        [3].0   // PV OUTPUT STATUS: SPARE
        [1].4   // PV OUTPUT STATUS: SPARE SOLENOID SV-372
        [3].4   // PV OUTPUT STATUS: SPARE
        [3].1   // PV OUTPUT STATUS: SPARE
        [4].12   // PV OUTPUT STATUS: SPARE
        [1].5   // PV OUTPUT STATUS: RETURN TO DRAIN XY-018
        [3].5   // PV OUTPUT STATUS: SPARE
        [4].13   // PV OUTPUT STATUS: SPARE
        [3].6   // PV OUTPUT STATUS: SPARE
        [3].10   // PV OUTPUT STATUS: SPARE
        [3].11   // PV OUTPUT STATUS: SPARE
        [1].1   // PV OUTPUT STATUS: AIR BLOW XV-008A
        [2].2   // PV OUTPUT STATUS: DRAIN TO WASTE NEUTRALIZATION XY-024
        [4].14   // PV OUTPUT STATUS: SPARE
        [1].6   // PV OUTPUT STATUS: ALARM HORN AH-376
        [4].9   // PV OUTPUT STATUS: SPARE
        [2].3   // PV OUTPUT STATUS: SPARE SOLENOID SV-410
        [5]   // PV OUTPUT STATUS: SCREEN 5
        [2].4   // PV OUTPUT STATUS: SPARE SOLENOID SV-412
        [1].10   // PV OUTPUT STATUS: CHEM #1 ENABLE XY-202
        [2].5   // PV OUTPUT STATUS: SPARE OUT-414
        [3].7   // PV OUTPUT STATUS: SPARE
        [2].6   // PV OUTPUT STATUS: SPARE OUT-416
        [4].15   // PV OUTPUT STATUS: SPARE
        [3].8   // PV OUTPUT STATUS: SPARE
        [6]   // PV OUTPUT STATUS: SCREEN 6
        [2].7   // PV OUTPUT STATUS: SPARE OUT-418
        [1].11   // PV OUTPUT STATUS: CHEM #2 ENABLE XY-302
        [3].9   // PV OUTPUT STATUS: SPARE
        [4].2   // PV OUTPUT STATUS: SPARE
        [1].7   // PV OUTPUT STATUS: HEATER ENABLE JY-004A
        [3].12   // PV OUTPUT STATUS: SPARE
        [4].3   // PV OUTPUT STATUS: SPARE
        [3].13   // PV OUTPUT STATUS: SPARE
        [1].12   // PV OUTPUT STATUS: CHEM #1 BLOCK XY-205
        [4]   // PV OUTPUT STATUS: SCREEN 4
        [7]   // PV OUTPUT STATUS: SCREEN 7
        [1].8   // PV OUTPUT STATUS: AIR BLOW BLOCK XY-008
        [4].0   // PV OUTPUT STATUS: SPARE
        [4].1   // PV OUTPUT STATUS: SPARE
        [1].9   // PV OUTPUT STATUS: SPARE OUT-384
        [2].8   // PV OUTPUT STATUS: SPARE
        [2]   // PV OUTPUT STATUS: SCREEN 2
        [3].14   // PV OUTPUT STATUS: SPARE
        [2].9   // PV OUTPUT STATUS: SPARE
        [1].13   // PV OUTPUT STATUS: CHEM #2 BLOCK XY-305
        [2].0   // PV OUTPUT STATUS: OVERFLOW TANK DRAIN XY-022
   PV_Output_Status_IND : INT[20,16] := ([1,6] := 1, [6,9] := 1, [6,11] := 1, [6,13] := 1, [7,0] := 1, [7,1] := 1, [7,2] := 1, [7,3] := 1, [7,4] := 1, [7,5] := 1);   // PV OUTPUT STATUS IND:
        [5,0]   // PV OUTPUT STATUS IND: SPARE
        [6,15]   // PV OUTPUT STATUS IND: SPARE
        [8,5]   // PV OUTPUT STATUS IND: SPARE
        [8,6]   // PV OUTPUT STATUS IND: SPARE
        [5,10]   // PV OUTPUT STATUS IND: SPARE
        [1,9]   // PV OUTPUT STATUS IND: SPARE OUT-384
        [9,8]   // PV OUTPUT STATUS IND: SPARE
        [4,12]   // PV OUTPUT STATUS IND: SPARE
        [5,9]   // PV OUTPUT STATUS IND: SPARE
        [9,9]   // PV OUTPUT STATUS IND: SPARE
        [8,7]   // PV OUTPUT STATUS IND: SPARE
        [6,1]   // PV OUTPUT STATUS IND: SPARE
        [5,11]   // PV OUTPUT STATUS IND: SPARE
        [5,12]   // PV OUTPUT STATUS IND: SPARE
        [7,4]   // PV OUTPUT STATUS IND: SPARE
        [1,0]   // PV OUTPUT STATUS IND: SPARE OUT-396
        [1,10]   // PV OUTPUT STATUS IND: CHEM #1 ENABLE XY-202
        [2,0]   // PV OUTPUT STATUS IND: OVERFLOW TANK DRAIN XY-022
        [1,11]   // PV OUTPUT STATUS IND: CHEM #2 ENABLE XY-302
        [2,10]   // PV OUTPUT STATUS IND: SPARE
        [8,8]   // PV OUTPUT STATUS IND: SPARE
        [7,11]   // PV OUTPUT STATUS IND: SPARE
        [5,13]   // PV OUTPUT STATUS IND: SPARE
        [6,0]   // PV OUTPUT STATUS IND: SPARE
        [1,12]   // PV OUTPUT STATUS IND: CHEM #1 BLOCK XY-205
        [8,9]   // PV OUTPUT STATUS IND: SPARE
        [3,4]   // PV OUTPUT STATUS IND: SPARE
        [5,14]   // PV OUTPUT STATUS IND: SPARE
        [6,2]   // PV OUTPUT STATUS IND: SPARE
        [1,13]   // PV OUTPUT STATUS IND: CHEM #2 BLOCK XY-305
        [1,14]   // PV OUTPUT STATUS IND: OVERFLOW TANK DRAIN PUMP XV-032
        [7,5]   // PV OUTPUT STATUS IND: SPARE
        [5,15]   // PV OUTPUT STATUS IND: SPARE
        [3,5]   // PV OUTPUT STATUS IND: SPARE
        [2,11]   // PV OUTPUT STATUS IND: SPARE
        [7,6]   // PV OUTPUT STATUS IND: SPARE
        [7,7]   // PV OUTPUT STATUS IND: SPARE
        [7,8]   // PV OUTPUT STATUS IND: SPARE
        [6,10]   // PV OUTPUT STATUS IND: SPARE
        [7,12]   // PV OUTPUT STATUS IND: SPARE
        [0,11]   // PV OUTPUT STATUS IND: NOT USED
        [0,12]   // PV OUTPUT STATUS IND: NOT USED
        [4,13]   // PV OUTPUT STATUS IND: SPARE
        [2,12]   // PV OUTPUT STATUS IND: SPARE
        [4,14]   // PV OUTPUT STATUS IND: SPARE
        [0,13]   // PV OUTPUT STATUS IND: NOT USED
        [9,0]   // PV OUTPUT STATUS IND: SPARE
        [4,15]   // PV OUTPUT STATUS IND: SPARE
        [6,3]   // PV OUTPUT STATUS IND: SPARE
        [6,11]   // PV OUTPUT STATUS IND: SPARE
        [1,15]   // PV OUTPUT STATUS IND: SPARE OUT-396
        [5,1]   // PV OUTPUT STATUS IND: SPARE
        [1,1]   // PV OUTPUT STATUS IND: AIR BLOW XV-008A
        [6,12]   // PV OUTPUT STATUS IND: SPARE
        [6,4]   // PV OUTPUT STATUS IND: SPARE
        [9,10]   // PV OUTPUT STATUS IND: SPARE
        [6,5]   // PV OUTPUT STATUS IND: SPARE
        [9,11]   // PV OUTPUT STATUS IND: SPARE
        [1,2]   // PV OUTPUT STATUS IND: SUPPLY PUMP CASING DRAIN XY-002
        [2,13]   // PV OUTPUT STATUS IND: SPARE
        [2,14]   // PV OUTPUT STATUS IND: SPARE
        [2,15]   // PV OUTPUT STATUS IND: SPARE
        [2,1]   // PV OUTPUT STATUS IND: LOW POINT DRAIN XY-023
        [2,2]   // PV OUTPUT STATUS IND: DRAIN TO WASTE NEUTRALIZATION XY-024
        [2,3]   // PV OUTPUT STATUS IND: SPARE SOLENOID SV-410
        [2,4]   // PV OUTPUT STATUS IND: SPARE SOLENOID SV-412
        [2,5]   // PV OUTPUT STATUS IND: SPARE OUT-414
        [2,6]   // PV OUTPUT STATUS IND: SPARE OUT-416
        [2,7]   // PV OUTPUT STATUS IND: SPARE OUT-418
        [7,13]   // PV OUTPUT STATUS IND: SPARE
        [7,9]   // PV OUTPUT STATUS IND: SPARE
        [7,14]   // PV OUTPUT STATUS IND: SPARE
        [0,14]   // PV OUTPUT STATUS IND: NOT USED
        [9,12]   // PV OUTPUT STATUS IND: SPARE
        [4,1]   // PV OUTPUT STATUS IND: SPARE
        [3,1]   // PV OUTPUT STATUS IND: SPARE
        [0,15]   // PV OUTPUT STATUS IND: NOT USED
        [7,15]   // PV OUTPUT STATUS IND: SPARE
        [6,6]   // PV OUTPUT STATUS IND: SPARE
        [6,7]   // PV OUTPUT STATUS IND: SPARE
        [8,0]   // PV OUTPUT STATUS IND: SPARE
        [1,3]   // PV OUTPUT STATUS IND: SUPPLY PUMP ENABLE JY-001A
        [3,6]   // PV OUTPUT STATUS IND: SPARE
        [9,13]   // PV OUTPUT STATUS IND: SPARE
        [9,14]   // PV OUTPUT STATUS IND: SPARE
        [0,1]   // PV OUTPUT STATUS IND: NOT USED
        [0,2]   // PV OUTPUT STATUS IND: NOT USED
        [0,3]   // PV OUTPUT STATUS IND: NOT USED
        [1,4]   // PV OUTPUT STATUS IND: SPARE SOLENOID SV-372
        [2,8]   // PV OUTPUT STATUS IND: SPARE
        [7,1]   // PV OUTPUT STATUS IND: SPARE
        [6,8]   // PV OUTPUT STATUS IND: SPARE
        [0,4]   // PV OUTPUT STATUS IND: NOT USED
        [4,2]   // PV OUTPUT STATUS IND: SPARE
        [1,5]   // PV OUTPUT STATUS IND: RETURN TO DRAIN XY-018
        [6,13]   // PV OUTPUT STATUS IND: SPARE
        [6,9]   // PV OUTPUT STATUS IND: SPARE
        [8,10]   // PV OUTPUT STATUS IND: SPARE
        [5,2]   // PV OUTPUT STATUS IND: SPARE
        [4,3]   // PV OUTPUT STATUS IND: SPARE
        [7,0]   // PV OUTPUT STATUS IND: SPARE
        [4,4]   // PV OUTPUT STATUS IND: SPARE
        [4,5]   // PV OUTPUT STATUS IND: SPARE
        [8,11]   // PV OUTPUT STATUS IND: SPARE
        [9,15]   // PV OUTPUT STATUS IND: SPARE
        [3,7]   // PV OUTPUT STATUS IND: SPARE
        [3,8]   // PV OUTPUT STATUS IND: SPARE
        [2,9]   // PV OUTPUT STATUS IND: SPARE
        [9,1]   // PV OUTPUT STATUS IND: SPARE
        [9,2]   // PV OUTPUT STATUS IND: SPARE
        [0,5]   // PV OUTPUT STATUS IND: NOT USED
        [3,9]   // PV OUTPUT STATUS IND: SPARE
        [4,6]   // PV OUTPUT STATUS IND: SPARE
        [5,3]   // PV OUTPUT STATUS IND: SPARE
        [0,6]   // PV OUTPUT STATUS IND: NOT USED
        [7,2]   // PV OUTPUT STATUS IND: SPARE
        [8,12]   // PV OUTPUT STATUS IND: SPARE
        [4,7]   // PV OUTPUT STATUS IND: SPARE
        [1,6]   // PV OUTPUT STATUS IND: ALARM HORN AH-376
        [1,7]   // PV OUTPUT STATUS IND: HEATER ENABLE JY-004A
        [3,0]   // PV OUTPUT STATUS IND: SPARE
        [0,7]   // PV OUTPUT STATUS IND: NOT USED
        [8,13]   // PV OUTPUT STATUS IND: SPARE
        [9,3]   // PV OUTPUT STATUS IND: SPARE
        [8,14]   // PV OUTPUT STATUS IND: SPARE
        [3,10]   // PV OUTPUT STATUS IND: SPARE
        [9,4]   // PV OUTPUT STATUS IND: SPARE
        [0,8]   // PV OUTPUT STATUS IND: NOT USED
        [8,15]   // PV OUTPUT STATUS IND: SPARE
        [9,5]   // PV OUTPUT STATUS IND: SPARE
        [9,6]   // PV OUTPUT STATUS IND: SPARE
        [0,0]   // PV OUTPUT STATUS IND: NOT USED
        [6,14]   // PV OUTPUT STATUS IND: SPARE
        [5,4]   // PV OUTPUT STATUS IND: SPARE
        [4,0]   // PV OUTPUT STATUS IND: SPARE
        [4,10]   // PV OUTPUT STATUS IND: SPARE
        [3,2]   // PV OUTPUT STATUS IND: SPARE
        [3,11]   // PV OUTPUT STATUS IND: SPARE
        [4,8]   // PV OUTPUT STATUS IND: SPARE
        [3,3]   // PV OUTPUT STATUS IND: SPARE
        [3,12]   // PV OUTPUT STATUS IND: SPARE
        [9,7]   // PV OUTPUT STATUS IND: SPARE
        [8,1]   // PV OUTPUT STATUS IND: SPARE
        [3,13]   // PV OUTPUT STATUS IND: SPARE
        [8,2]   // PV OUTPUT STATUS IND: SPARE
        [4,11]   // PV OUTPUT STATUS IND: SPARE
        [4,9]   // PV OUTPUT STATUS IND: SPARE
        [1,8]   // PV OUTPUT STATUS IND: AIR BLOW BLOCK XY-008
        [3,14]   // PV OUTPUT STATUS IND: SPARE
        [0,9]   // PV OUTPUT STATUS IND: NOT USED
        [5,5]   // PV OUTPUT STATUS IND: SPARE
        [5,6]   // PV OUTPUT STATUS IND: SPARE
        [5,7]   // PV OUTPUT STATUS IND: SPARE
        [7,10]   // PV OUTPUT STATUS IND: SPARE
        [0,10]   // PV OUTPUT STATUS IND: NOT USED
        [8,3]   // PV OUTPUT STATUS IND: SPARE
        [5,8]   // PV OUTPUT STATUS IND: SPARE
        [7,3]   // PV OUTPUT STATUS IND: SPARE
        [8,4]   // PV OUTPUT STATUS IND: SPARE
        [3,15]   // PV OUTPUT STATUS IND: SPARE
   PV_Rename_Recipe_Name : STRING := 'RECIPE #35';   // PANELVIEW RENAME RECIPE NAME
   PV_Status_Bit : BOOL := 1;   // SYSTEM BIT
   PV_Step_Time : DINT;   // PANELVIEW DISPLAY STEP TIME
   pv_step_time_minutes : DINT;   // PANELVIEW DISPLAY STEP TIME MINUTES
   pv_step_time_seconds : DINT;   // PANELVIEW DISPLAY STEP TIME SECONDS
   PV_Visibility : DINT[4] := ([0] := -1981313, [2] := 32, [3] := 20);   // HMI VISIBILITY CONTROL BITS 0 = AVAILABLE / 1 = GREY
        [2].2   // PLC CLOCK UPDATE PUSHBUTTONS VISIBILITY 0 = AVAILABLE / 1 = GREY
        [0].15   // SPARE PUSHBUTTONS VISIBILITY 0 = AVAILABLE / 1 = GREY
        [0].2   // HOLD PUSHBUTTON VISIBILITY 0 = AVAILABLE / 1 = GREY
        [1].12   // SPARE PUSHBUTTONS VISIBILITY 0 = AVAILABLE / 1 = GREY
        [2].5   // SUPPLY TEMPERATURE PID IN MANUAL/AUTO PUSHBUTTONS VISIBILITY 0 = AVAILABLE / 1 = GREY
        [3].12   // SPARE PUSHBUTTON VISIBILITY
        [2].3   // COPY RECIPES PUSHBUTTON VISIBILITY 0 = AVAILABLE 1 = GREY
        [0].3   // SPARE PUSHBUTTONS VISIBILITY 0 = AVAILABLE / 1 = GREY
        [3].13   // SPARE PUSHBUTTON VISIBILITY
        [0].4   // ABORT PUSHBUTTON VISIBILITY 0 = AVAILABLE / 1 = GREY
        [0]   // HMI VISIBILITY CONTROL BITS FOR CONTROLLER SCREEN
        [1].13   // SPARE PUSHBUTTONS VISIBILITY 0 = AVAILABLE / 1 = GREY
        [1].14   // SPARE PUSHBUTTONS VISIBILITY 0 = AVAILABLE / 1 = GREY
        [0].5   // STEP PUSHBUTTON VISIBILITY 0 = AVAILABLE / 1 = GREY
        [1].15   // SPARE PUSHBUTTONS VISIBILITY 0 = AVAILABLE / 1 = GREY
        [0].0   // START PUSHBUTTON VISIBILITY 0 = AVAILABLE / 1 = GREY
        [3].14   // SPARE PUSHBUTTON VISIBILITY
        [0].1   // STOP PUSHBUTTON VISIBILITY 0 = AVAILABLE / 1 = GREY
        [3].15   // SPARE PUSHBUTTON VISIBILITY
        [2].4   // SPARE PUSHBUTTONS VISIBILITY 0 = AVAILABLE / 1 = GREY
        [0].6   // ALL AUTO PUSHBUTTON VISIBILITY 0 = AVAILABLE / 1 = GREY
        [3].2   // SPARE PUSHBUTTON VISIBILITY
        [3].3   // SPARE PUSHBUTTON VISIBILITY
        [2].6   // SPARE PUSHBUTTONS VISIBILITY 0 = AVAILABLE / 1 = GREY
        [3].4   // SPARE PUSHBUTTON VISIBILITY
        [0].7   // RECIPE PUSHBUTTON VISIBILITY 0 = AVAILABLE / 1 = GREY
        [0].10   // SPARE PUSHBUTTONS VISIBILITY 0 = AVAILABLE / 1 = GREY
        [2].7   // SPARE PUSHBUTTONS VISIBILITY 0 = AVAILABLE / 1 = GREY
        [0].8   // PRINT PUSHBUTTONS VISIBILITY 0 = AVAILABLE / 1 = GREY
        [3].5   // SPARE PUSHBUTTON VISIBILITY
        [2].8   // SPARE PUSHBUTTONS VISIBILITY 0 = AVAILABLE / 1 = GREY
        [3].6   // SPARE PUSHBUTTON VISIBILITY
        [3].7   // SPARE PUSHBUTTON VISIBILITY
        [0].11   // SPARE PUSHBUTTONS VISIBILITY 0 = AVAILABLE / 1 = GREY
        [2]   // HMI VISIBILITY CONTROL BITS FOR RECIPE EDIT SCREENS
        [3].8   // SPARE PUSHBUTTON VISIBILITY
        [0].12   // SPARE PUSHBUTTONS VISIBILITY 0 = AVAILABLE / 1 = GREY
        [1].2   // DRAIN PUSHBUTTONS VISIBILITY 0 = AVAILABLE / 1 = GREY
        [3].9   // SPARE PUSHBUTTON VISIBILITY
        [0].9   // HEATER MOA PUSHBUTTON VISIBILITY 0 = AVAILABLE / 1 = GREY
        [0].13   // SPARE PUSHBUTTONS VISIBILITY 0 = AVAILABLE / 1 = GREY
        [1]   // HMI VISIBILITY CONTROL BITS FOR UTILITY SCREEN
        [1].3   // CHEM #1 ENABLE PUSHBUTTONS VISIBILITY 0 = AVAILABLE / 1 = GREY
        [2].0   // INSERT STEP PUSHBUTTONS VISIBILITY 0 = AVAILABLE / 1 = GREY
        [0].14   // SPARE PUSHBUTTONS VISIBILITY 0 = AVAILABLE / 1 = GREY
        [2].9   // SPARE PUSHBUTTONS VISIBILITY 0 = AVAILABLE / 1 = GREY
        [1].0   // PW ENABLE PUSHBUTTONS VISIBILITY 0 = AVAILABLE / 1 = GREY
        [1].4   // CHEM #2 ENABLE PUSHBUTTONS VISIBILITY 0 = AVAILABLE / 1 = GREY
        [3]   // PLC CLOCK UPDATE PUSHBUTTONS VISIBILITY DURATION
        [1].5   // SPARE PUSHBUTTONS VISIBILITY 0 = AVAILABLE / 1 = GREY
        [1].1   // WFI ENABLE PUSHBUTTONS VISIBILITY 0 = AVAILABLE / 1 = GREY
        [1].6   // SPARE PUSHBUTTONS VISIBILITY 0 = AVAILABLE / 1 = GREY
        [3].0   // SPARE PUSHBUTTON VISIBILITY
        [3].1   // SPARE PUSHBUTTON VISIBILITY
        [1].7   // SPARE PUSHBUTTONS VISIBILITY 0 = AVAILABLE / 1 = GREY
        [2].1   // DELETE STEP PUSHBUTTONS VISIBILITY 0 = AVAILABLE / 1 = GREY
        [1].8   // SPARE PUSHBUTTONS VISIBILITY 0 = AVAILABLE / 1 = GREY
        [2].10   // SPARE PUSHBUTTONS VISIBILITY 0 = AVAILABLE / 1 = GREY
        [3].10   // SPARE PUSHBUTTON VISIBILITY
        [1].10   // SPARE PUSHBUTTONS VISIBILITY 0 = AVAILABLE / 1 = GREY
        [2].11   // SPARE PUSHBUTTONS VISIBILITY 0 = AVAILABLE / 1 = GREY
        [2].12   // SPARE PUSHBUTTONS VISIBILITY 0 = AVAILABLE / 1 = GREY
        [1].9   // SPARE PUSHBUTTONS VISIBILITY 0 = AVAILABLE / 1 = GREY
        [3].11   // SPARE PUSHBUTTON VISIBILITY
        [1].11   // SPARE PUSHBUTTONS VISIBILITY 0 = AVAILABLE / 1 = GREY
        [2].13   // SPARE PUSHBUTTONS VISIBILITY 0 = AVAILABLE / 1 = GREY
        [2].14   // SPARE PUSHBUTTONS VISIBILITY 0 = AVAILABLE / 1 = GREY
        [2].15   // SPARE PUSHBUTTONS VISIBILITY 0 = AVAILABLE / 1 = GREY
   Recipe : RECIPE[41] := ([0].OpCode[1] := 4, [0].OpCode[2] := 8, [0].OpCode[3] := 9, [0].OpCode[4] := 5, [0].OpCode[5] := 4, [0].OpCode[6] := 7, [0].OpCode[7] := 10, [0].OpCode[8] := 13, [0].OpCode[9] := 16, [0].OpCode[10] := 20, [0].OpCode[11] := 5, [0].OpCode[12] := 4, [0].OpCode[13] := 11, [0].OpCode[14] := 13, [0].OpCode[15] := 16, [0].OpCode[16] := 14, [0].OpCode[17] := 17, [0].OpCode[18] := 18, [0].OpCode[19] := 2, [0].OpCode[20] := 1, [0].StepTime[1] := 10, [0].StepTime[2] := 10, [0].StepTime[3] := 10, [0].StepTime[4] := 10, [0].StepTime[5] := 10, [0].StepTime[6] := 10, [0].StepTime[7] := 10, [0].StepTime[8] := 10, [0].StepTime[9] := 10, [0].StepTime[10] := 10, [0].StepTime[11] := 10, [0].StepTime[12] := 10, [0].StepTime[13] := 10, [0].StepTime[14] := 10, [0].StepTime[15] := 10, [0].StepTime[16] := 10, [0].StepTime[17] := 10, [0].StepTime[18] := 10, [0].StepTime[19] := 10, [0].StepTime[20] := 10, [0].Setpoint[1] := 55.0, [0].Setpoint[2] := 65.0, [0].Setpoint[3] := 60.0, [0].Setpoint[4] := 45.0, [0].Setpoint[5] := 65.0, [0].Setpoint[7] := 53.0, [0].Setpoint[8] := 63.0, [0].Setpoint[9] := 57.0, [0].Setpoint[10] := 43.0, [0].Setpoint[11] := 63.0, [0].Setpoint[13] := 85.0, [0].Setpoint[14] := 300.0, [0].Setpoint[15] := 900.0, [0].Setpoint[17] := 15.0, [0].Setpoint[18] := 14.0, [0].Setpoint[19] := 15.0, [0].Setpoint[20] := 45.0, [0].Setpoint[21] := 5.0, [0].Setpoint[22] := 15.0, [0].Setpoint[23] := 300.0,
        [0].Setpoint[25] := 10.0, [0].Setpoint[26] := 9.0, [0].Setpoint[27] := 10.0, [0].Setpoint[28] := 50.0, [0].Setpoint[29] := 3.0, [0].Setpoint[30] := 17.0, [0].Setpoint[31] := 300.0, [0].Setpoint[33] := 2.0, [0].Setpoint[34] := 900.0, [0].Setpoint[37] := 35.0, [0].Setpoint[41] := 5.0, [0].Setpoint[42] := 50.0, [0].Setpoint[43] := 5.0, [0].Setpoint[44] := 60.0, [0].Setpoint[45] := 50.0, [0].Setpoint[47] := 15.0, [0].Setpoint[49] := 180.0, [0].Setpoint[50] := 180.0, [0].Setpoint[52] := 30.0, [0].Setpoint[53] := 5.0, [0].Setpoint[54] := 5.0, [0].Setpoint[55] := 3.0, [0].Setpoint[57] := 300.0, [0].Name := 'FAT TEST RECIPE', [1].OpCode[1] := 4, [1].OpCode[2] := 9, [1].OpCode[3] := 5, [1].OpCode[4] := 2, [1].OpCode[5] := 4, [1].OpCode[6] := 10, [1].OpCode[7] := 17, [1].OpCode[8] := 5, [1].OpCode[9] := 2, [1].OpCode[10] := 4, [1].OpCode[11] := 16, [1].OpCode[12] := 5, [1].OpCode[13] := 2, [1].OpCode[14] := 4, [1].OpCode[15] := 11, [1].OpCode[16] := 17, [1].OpCode[17] := 5, [1].OpCode[18] := 2, [1].OpCode[19] := 4, [1].OpCode[20] := 16, [1].OpCode[21] := 5, [1].OpCode[22] := 2, [1].OpCode[23] := 4, [1].OpCode[24] := 16, [1].OpCode[25] := 5, [1].OpCode[26] := 2, [1].OpCode[27] := 4, [1].OpCode[28] := 14, [1].OpCode[29] := 5, [1].OpCode[30] := 2, [1].OpCode[31] := 1, [1].StepTime[1] := 1, [1].StepTime[2] := 120, [1].StepTime[3] := 1, [1].StepTime[4] := 10, [1].StepTime[5] := 1,
        [1].StepTime[6] := 150, [1].StepTime[7] := 5, [1].StepTime[8] := 1, [1].StepTime[9] := 10, [1].StepTime[10] := 1, [1].StepTime[11] := 50, [1].StepTime[12] := 1, [1].StepTime[13] := 10, [1].StepTime[14] := 1, [1].StepTime[15] := 150, [1].StepTime[16] := 5, [1].StepTime[17] := 1, [1].StepTime[18] := 10, [1].StepTime[19] := 1, [1].StepTime[20] := 50, [1].StepTime[21] := 1, [1].StepTime[22] := 10, [1].StepTime[23] := 1, [1].StepTime[24] := 50, [1].StepTime[25] := 1, [1].StepTime[26] := 10, [1].StepTime[27] := 1, [1].StepTime[28] := 50, [1].StepTime[29] := 1, [1].StepTime[30] := 10, [1].StepTime[31] := 1, [1].Setpoint[1] := 55.0, [1].Setpoint[2] := 65.0, [1].Setpoint[3] := 60.0, [1].Setpoint[4] := 45.0, [1].Setpoint[5] := 65.0, [1].Setpoint[7] := 53.0, [1].Setpoint[8] := 63.0, [1].Setpoint[9] := 57.0, [1].Setpoint[10] := 43.0, [1].Setpoint[11] := 63.0, [1].Setpoint[13] := 85.0, [1].Setpoint[14] := 300.0, [1].Setpoint[15] := 900.0, [1].Setpoint[17] := 15.0, [1].Setpoint[18] := 14.0, [1].Setpoint[19] := 15.0, [1].Setpoint[20] := 45.0, [1].Setpoint[21] := 5.0, [1].Setpoint[22] := 15.0, [1].Setpoint[23] := 300.0, [1].Setpoint[25] := 10.0, [1].Setpoint[26] := 9.0, [1].Setpoint[27] := 10.0, [1].Setpoint[28] := 50.0, [1].Setpoint[29] := 3.0, [1].Setpoint[30] := 17.0, [1].Setpoint[31] := 300.0, [1].Setpoint[33] := 2.0, [1].Setpoint[34] := 900.0, [1].Setpoint[37] := 35.0, [1].Setpoint[41] := 5.0, [1].Setpoint[42] := 50.0, [1].Setpoint[43] := 5.0, [1].Setpoint[44] := 60.0,
        [1].Setpoint[45] := 50.0, [1].Setpoint[47] := 15.0, [1].Setpoint[49] := 180.0, [1].Setpoint[50] := 180.0, [1].Setpoint[52] := 30.0, [1].Setpoint[53] := 5.0, [1].Setpoint[54] := 5.0, [1].Setpoint[55] := 3.0, [1].Setpoint[56] := 1.0, [1].Setpoint[57] := 300.0, [1].Name := 'WASH CYCLE', [2].Setpoint[1] := 55.0, [2].Setpoint[2] := 65.0, [2].Setpoint[3] := 60.0, [2].Setpoint[4] := 45.0, [2].Setpoint[5] := 65.0, [2].Setpoint[7] := 53.0, [2].Setpoint[8] := 63.0, [2].Setpoint[9] := 57.0, [2].Setpoint[10] := 43.0, [2].Setpoint[11] := 63.0, [2].Setpoint[13] := 85.0, [2].Setpoint[14] := 300.0, [2].Setpoint[15] := 900.0, [2].Setpoint[17] := 15.0, [2].Setpoint[18] := 14.0, [2].Setpoint[19] := 15.0, [2].Setpoint[20] := 45.0, [2].Setpoint[21] := 5.0, [2].Setpoint[22] := 15.0, [2].Setpoint[23] := 300.0, [2].Setpoint[25] := 10.0, [2].Setpoint[26] := 9.0, [2].Setpoint[27] := 10.0, [2].Setpoint[28] := 50.0, [2].Setpoint[29] := 3.0, [2].Setpoint[30] := 17.0, [2].Setpoint[31] := 300.0, [2].Setpoint[33] := 2.0, [2].Setpoint[34] := 900.0, [2].Setpoint[37] := 35.0, [2].Setpoint[41] := 5.0, [2].Setpoint[42] := 50.0, [2].Setpoint[43] := 5.0, [2].Setpoint[44] := 60.0, [2].Setpoint[45] := 50.0, [2].Setpoint[47] := 15.0, [2].Setpoint[49] := 180.0, [2].Setpoint[50] := 180.0, [2].Setpoint[52] := 30.0, [2].Setpoint[53] := 5.0, [2].Setpoint[54] := 5.0, [2].Setpoint[55] := 3.0, [2].Setpoint[57] := 300.0, [2].Name := 'RECIPE #2', [3].Setpoint[1] := 55.0, [3].Setpoint[2] := 65.0, [3].Setpoint[3] := 60.0, [3].Setpoint[4] := 45.0, [3].Setpoint[5] := 65.0,
        [3].Setpoint[7] := 53.0, [3].Setpoint[8] := 63.0, [3].Setpoint[9] := 57.0, [3].Setpoint[10] := 43.0, [3].Setpoint[11] := 63.0, [3].Setpoint[13] := 85.0, [3].Setpoint[14] := 300.0, [3].Setpoint[15] := 900.0, [3].Setpoint[17] := 15.0, [3].Setpoint[18] := 14.0, [3].Setpoint[19] := 15.0, [3].Setpoint[20] := 45.0, [3].Setpoint[21] := 5.0, [3].Setpoint[22] := 15.0, [3].Setpoint[23] := 300.0, [3].Setpoint[25] := 10.0, [3].Setpoint[26] := 9.0, [3].Setpoint[27] := 10.0, [3].Setpoint[28] := 50.0, [3].Setpoint[29] := 3.0, [3].Setpoint[30] := 17.0, [3].Setpoint[31] := 300.0, [3].Setpoint[33] := 2.0, [3].Setpoint[34] := 900.0, [3].Setpoint[37] := 35.0, [3].Setpoint[41] := 5.0, [3].Setpoint[42] := 50.0, [3].Setpoint[43] := 5.0, [3].Setpoint[44] := 60.0, [3].Setpoint[45] := 50.0, [3].Setpoint[47] := 15.0, [3].Setpoint[49] := 180.0, [3].Setpoint[50] := 180.0, [3].Setpoint[52] := 30.0, [3].Setpoint[53] := 5.0, [3].Setpoint[54] := 5.0, [3].Setpoint[55] := 3.0, [3].Setpoint[57] := 300.0, [3].Name := 'RECIPE #3', [4].Setpoint[1] := 55.0, [4].Setpoint[2] := 65.0, [4].Setpoint[3] := 60.0, [4].Setpoint[4] := 45.0, [4].Setpoint[5] := 65.0, [4].Setpoint[7] := 53.0, [4].Setpoint[8] := 63.0, [4].Setpoint[9] := 57.0, [4].Setpoint[10] := 43.0, [4].Setpoint[11] := 63.0, [4].Setpoint[13] := 85.0, [4].Setpoint[14] := 300.0, [4].Setpoint[15] := 900.0, [4].Setpoint[17] := 15.0, [4].Setpoint[18] := 14.0, [4].Setpoint[19] := 15.0, [4].Setpoint[20] := 45.0, [4].Setpoint[21] := 5.0, [4].Setpoint[22] := 15.0, [4].Setpoint[23] := 300.0, [4].Setpoint[25] := 10.0,
        [4].Setpoint[26] := 9.0, [4].Setpoint[27] := 10.0, [4].Setpoint[28] := 50.0, [4].Setpoint[29] := 3.0, [4].Setpoint[30] := 17.0, [4].Setpoint[31] := 300.0, [4].Setpoint[33] := 2.0, [4].Setpoint[34] := 900.0, [4].Setpoint[37] := 35.0, [4].Setpoint[41] := 5.0, [4].Setpoint[42] := 50.0, [4].Setpoint[43] := 5.0, [4].Setpoint[44] := 60.0, [4].Setpoint[45] := 50.0, [4].Setpoint[47] := 15.0, [4].Setpoint[49] := 180.0, [4].Setpoint[50] := 180.0, [4].Setpoint[52] := 30.0, [4].Setpoint[53] := 5.0, [4].Setpoint[54] := 5.0, [4].Setpoint[55] := 3.0, [4].Setpoint[57] := 300.0, [4].Name := 'RECIPE #4', [5].Setpoint[1] := 55.0, [5].Setpoint[2] := 65.0, [5].Setpoint[3] := 60.0, [5].Setpoint[4] := 45.0, [5].Setpoint[5] := 65.0, [5].Setpoint[7] := 53.0, [5].Setpoint[8] := 63.0, [5].Setpoint[9] := 57.0, [5].Setpoint[10] := 43.0, [5].Setpoint[11] := 63.0, [5].Setpoint[13] := 85.0, [5].Setpoint[14] := 300.0, [5].Setpoint[15] := 900.0, [5].Setpoint[17] := 15.0, [5].Setpoint[18] := 14.0, [5].Setpoint[19] := 15.0, [5].Setpoint[20] := 45.0, [5].Setpoint[21] := 5.0, [5].Setpoint[22] := 15.0, [5].Setpoint[23] := 300.0, [5].Setpoint[25] := 10.0, [5].Setpoint[26] := 9.0, [5].Setpoint[27] := 10.0, [5].Setpoint[28] := 50.0, [5].Setpoint[29] := 3.0, [5].Setpoint[30] := 17.0, [5].Setpoint[31] := 300.0, [5].Setpoint[33] := 2.0, [5].Setpoint[34] := 900.0, [5].Setpoint[37] := 35.0, [5].Setpoint[41] := 5.0, [5].Setpoint[42] := 50.0, [5].Setpoint[43] := 5.0, [5].Setpoint[44] := 60.0, [5].Setpoint[45] := 50.0, [5].Setpoint[47] := 15.0, [5].Setpoint[49] := 180.0,
        [5].Setpoint[50] := 180.0, [5].Setpoint[52] := 30.0, [5].Setpoint[53] := 5.0, [5].Setpoint[54] := 5.0, [5].Setpoint[55] := 3.0, [5].Setpoint[57] := 300.0, [5].Name := 'RECIPE #5', [6].Setpoint[1] := 55.0, [6].Setpoint[2] := 65.0, [6].Setpoint[3] := 60.0, [6].Setpoint[4] := 45.0, [6].Setpoint[5] := 65.0, [6].Setpoint[7] := 53.0, [6].Setpoint[8] := 63.0, [6].Setpoint[9] := 57.0, [6].Setpoint[10] := 43.0, [6].Setpoint[11] := 63.0, [6].Setpoint[13] := 85.0, [6].Setpoint[14] := 300.0, [6].Setpoint[15] := 900.0, [6].Setpoint[17] := 15.0, [6].Setpoint[18] := 14.0, [6].Setpoint[19] := 15.0, [6].Setpoint[20] := 45.0, [6].Setpoint[21] := 5.0, [6].Setpoint[22] := 15.0, [6].Setpoint[23] := 300.0, [6].Setpoint[25] := 10.0, [6].Setpoint[26] := 9.0, [6].Setpoint[27] := 10.0, [6].Setpoint[28] := 50.0, [6].Setpoint[29] := 3.0, [6].Setpoint[30] := 17.0, [6].Setpoint[31] := 300.0, [6].Setpoint[33] := 2.0, [6].Setpoint[34] := 900.0, [6].Setpoint[37] := 35.0, [6].Setpoint[41] := 5.0, [6].Setpoint[42] := 50.0, [6].Setpoint[43] := 5.0, [6].Setpoint[44] := 60.0, [6].Setpoint[45] := 50.0, [6].Setpoint[47] := 15.0, [6].Setpoint[49] := 180.0, [6].Setpoint[50] := 180.0, [6].Setpoint[52] := 30.0, [6].Setpoint[53] := 5.0, [6].Setpoint[54] := 5.0, [6].Setpoint[55] := 3.0, [6].Setpoint[57] := 300.0, [6].Name := 'RECIPE #6', [7].Setpoint[1] := 55.0, [7].Setpoint[2] := 65.0, [7].Setpoint[3] := 60.0, [7].Setpoint[4] := 45.0, [7].Setpoint[5] := 65.0, [7].Setpoint[7] := 53.0, [7].Setpoint[8] := 63.0, [7].Setpoint[9] := 57.0, [7].Setpoint[10] := 43.0,
        [7].Setpoint[11] := 63.0, [7].Setpoint[13] := 85.0, [7].Setpoint[14] := 300.0, [7].Setpoint[15] := 900.0, [7].Setpoint[17] := 15.0, [7].Setpoint[18] := 14.0, [7].Setpoint[19] := 15.0, [7].Setpoint[20] := 45.0, [7].Setpoint[21] := 5.0, [7].Setpoint[22] := 15.0, [7].Setpoint[23] := 300.0, [7].Setpoint[25] := 10.0, [7].Setpoint[26] := 9.0, [7].Setpoint[27] := 10.0, [7].Setpoint[28] := 50.0, [7].Setpoint[29] := 3.0, [7].Setpoint[30] := 17.0, [7].Setpoint[31] := 300.0, [7].Setpoint[33] := 2.0, [7].Setpoint[34] := 900.0, [7].Setpoint[37] := 35.0, [7].Setpoint[41] := 5.0, [7].Setpoint[42] := 50.0, [7].Setpoint[43] := 5.0, [7].Setpoint[44] := 60.0, [7].Setpoint[45] := 50.0, [7].Setpoint[47] := 15.0, [7].Setpoint[49] := 180.0, [7].Setpoint[50] := 180.0, [7].Setpoint[52] := 30.0, [7].Setpoint[53] := 5.0, [7].Setpoint[54] := 5.0, [7].Setpoint[55] := 3.0, [7].Setpoint[57] := 300.0, [7].Name := 'RECIPE #7', [8].Setpoint[1] := 55.0, [8].Setpoint[2] := 65.0, [8].Setpoint[3] := 60.0, [8].Setpoint[4] := 45.0, [8].Setpoint[5] := 65.0, [8].Setpoint[7] := 53.0, [8].Setpoint[8] := 63.0, [8].Setpoint[9] := 57.0, [8].Setpoint[10] := 43.0, [8].Setpoint[11] := 63.0, [8].Setpoint[13] := 85.0, [8].Setpoint[14] := 300.0, [8].Setpoint[15] := 900.0, [8].Setpoint[17] := 15.0, [8].Setpoint[18] := 14.0, [8].Setpoint[19] := 15.0, [8].Setpoint[20] := 45.0, [8].Setpoint[21] := 5.0, [8].Setpoint[22] := 15.0, [8].Setpoint[23] := 300.0, [8].Setpoint[25] := 10.0, [8].Setpoint[26] := 9.0, [8].Setpoint[27] := 10.0, [8].Setpoint[28] := 50.0, [8].Setpoint[29] := 3.0,
        [8].Setpoint[30] := 17.0, [8].Setpoint[31] := 300.0, [8].Setpoint[33] := 2.0, [8].Setpoint[34] := 900.0, [8].Setpoint[37] := 35.0, [8].Setpoint[41] := 5.0, [8].Setpoint[42] := 50.0, [8].Setpoint[43] := 5.0, [8].Setpoint[44] := 60.0, [8].Setpoint[45] := 50.0, [8].Setpoint[47] := 15.0, [8].Setpoint[49] := 180.0, [8].Setpoint[50] := 180.0, [8].Setpoint[52] := 30.0, [8].Setpoint[53] := 5.0, [8].Setpoint[54] := 5.0, [8].Setpoint[55] := 3.0, [8].Setpoint[57] := 300.0, [8].Name := 'RECIPE #8', [9].Setpoint[1] := 55.0, [9].Setpoint[2] := 65.0, [9].Setpoint[3] := 60.0, [9].Setpoint[4] := 45.0, [9].Setpoint[5] := 65.0, [9].Setpoint[7] := 53.0, [9].Setpoint[8] := 63.0, [9].Setpoint[9] := 57.0, [9].Setpoint[10] := 43.0, [9].Setpoint[11] := 63.0, [9].Setpoint[13] := 85.0, [9].Setpoint[14] := 300.0, [9].Setpoint[15] := 900.0, [9].Setpoint[17] := 15.0, [9].Setpoint[18] := 14.0, [9].Setpoint[19] := 15.0, [9].Setpoint[20] := 45.0, [9].Setpoint[21] := 5.0, [9].Setpoint[22] := 15.0, [9].Setpoint[23] := 300.0, [9].Setpoint[25] := 10.0, [9].Setpoint[26] := 9.0, [9].Setpoint[27] := 10.0, [9].Setpoint[28] := 50.0, [9].Setpoint[29] := 3.0, [9].Setpoint[30] := 17.0, [9].Setpoint[31] := 300.0, [9].Setpoint[33] := 2.0, [9].Setpoint[34] := 900.0, [9].Setpoint[37] := 35.0, [9].Setpoint[41] := 5.0, [9].Setpoint[42] := 50.0, [9].Setpoint[43] := 5.0, [9].Setpoint[44] := 60.0, [9].Setpoint[45] := 50.0, [9].Setpoint[47] := 15.0, [9].Setpoint[49] := 180.0, [9].Setpoint[50] := 180.0, [9].Setpoint[52] := 30.0, [9].Setpoint[53] := 5.0, [9].Setpoint[54] := 5.0,
